(* IEC 61131-3 sources: plc-st-coding-agent/progress/evidence/f14_v10_full_20261113/jobs/codex_deepseek-v4pro (part 2) *)

(* ---- public-medium-05.candidate_02.st ---- *)
FUNCTION_BLOCK ProductionLineControl
(*
ENGINEERING_CONTRACT
MotorForward (PUB006/PUB007): manual ForwardButton iff not ReverseButton; auto hold while AutoStep=1 or AutoStep=3; deactivate at destination sensor B/C or on manual release/non-auto; simultaneous Forward/Reverse gives no motion.
MotorReverse (PUB004): manual ReverseButton iff not ForwardButton.
CompletionLight (PUB008): auto activate when C is reached and SensorC and ButtonC are TRUE, including same-scan arrival; retain while SensorC TRUE; reset only when SensorC FALSE.
AutoStep retains sequence state across scans; BOOL buttons are level-gated, no unstated edges.
*)
(* CONTRACT_RULES [] *)
VAR_INPUT
    Mode : BOOL;
    ForwardButton : BOOL;
    ReverseButton : BOOL;
    SensorA : BOOL;
    SensorB : BOOL;
    SensorC : BOOL;
    ButtonA : BOOL;
    ButtonB : BOOL;
    ButtonC : BOOL;
END_VAR
VAR_OUTPUT
    MotorForward : BOOL;
    MotorReverse : BOOL;
    CompletionLight : BOOL;
END_VAR
VAR
    AutoStep : INT := 0;
END_VAR

MotorForward := FALSE;
MotorReverse := FALSE;

IF NOT SensorC THEN
    CompletionLight := FALSE;
END_IF;

IF Mode THEN
    CASE AutoStep OF
        0:
            IF SensorA AND ButtonA THEN
                AutoStep := 1;
                MotorForward := TRUE;
            END_IF;

        1:
            IF SensorB THEN
                IF ButtonB THEN
                    AutoStep := 3;
                    MotorForward := TRUE;
                ELSE
                    AutoStep := 2;
                END_IF;
            ELSE
                MotorForward := TRUE;
            END_IF;

        2:
            IF ButtonB THEN
                AutoStep := 3;
                MotorForward := TRUE;
            END_IF;

        3:
            IF SensorC THEN
                AutoStep := 4;
                IF ButtonC THEN
                    CompletionLight := TRUE;
                END_IF;
            ELSE
                MotorForward := TRUE;
            END_IF;

        4:
            IF SensorC AND ButtonC THEN
                CompletionLight := TRUE;
            END_IF;
            IF NOT SensorC THEN
                AutoStep := 0;
            END_IF;
    END_CASE;
ELSE
    MotorForward := ForwardButton AND NOT ReverseButton;
    MotorReverse := ReverseButton AND NOT ForwardButton;
END_IF;
END_FUNCTION_BLOCK

(* ---- public-medium-05.candidate_03.st ---- *)
FUNCTION_BLOCK ProductionLineControl
(*
ENGINEERING_CONTRACT
MotorForward (PUB006/PUB007): manual ForwardButton iff not ReverseButton; auto hold while AutoStep=1 or AutoStep=3; deactivate at destination sensor B/C or on manual release/non-auto; simultaneous Forward/Reverse gives no motion.
MotorReverse (PUB004): manual ReverseButton iff not ForwardButton.
CompletionLight (PUB008): auto activate when C is reached and SensorC and ButtonC are TRUE, including same-scan arrival; retain while SensorC TRUE; reset only when SensorC FALSE.
AutoStep retains sequence state across scans; BOOL buttons are level-gated, no unstated edges.
*)
(* CONTRACT_RULES [] *)
VAR_INPUT
    Mode : BOOL;
    ForwardButton : BOOL;
    ReverseButton : BOOL;
    SensorA : BOOL;
    SensorB : BOOL;
    SensorC : BOOL;
    ButtonA : BOOL;
    ButtonB : BOOL;
    ButtonC : BOOL;
END_VAR
VAR_OUTPUT
    MotorForward : BOOL;
    MotorReverse : BOOL;
    CompletionLight : BOOL;
END_VAR
VAR
    AutoStep : INT := 0;
END_VAR

MotorForward := FALSE;
MotorReverse := FALSE;

IF NOT SensorC THEN
    CompletionLight := FALSE;
END_IF;

IF Mode THEN
    CASE AutoStep OF
        0:
            IF SensorA AND ButtonA THEN
                AutoStep := 1;
                MotorForward := TRUE;
            END_IF;

        1:
            IF SensorB THEN
                IF ButtonB THEN
                    AutoStep := 3;
                    MotorForward := TRUE;
                ELSE
                    AutoStep := 2;
                END_IF;
            ELSE
                MotorForward := TRUE;
            END_IF;

        2:
            IF ButtonB THEN
                AutoStep := 3;
                MotorForward := TRUE;
            END_IF;

        3:
            IF SensorC THEN
                AutoStep := 4;
                IF ButtonC THEN
                    CompletionLight := TRUE;
                END_IF;
            ELSE
                MotorForward := TRUE;
            END_IF;

        4:
            IF SensorC AND (CompletionLight OR ButtonC) THEN
                CompletionLight := TRUE;
            END_IF;
            IF NOT SensorC THEN
                AutoStep := 0;
            END_IF;
    END_CASE;
ELSE
    MotorForward := ForwardButton AND NOT ReverseButton;
    MotorReverse := ReverseButton AND NOT ForwardButton;
END_IF;
END_FUNCTION_BLOCK

(* ---- public-medium-05.raw_candidate_01.st ---- *)
FUNCTION_BLOCK ProductionLineControl
(*
ENGINEERING_CONTRACT
MotorForward (PUB001/PUB002/PUB003): activate manual ForwardButton or auto transfer state; hold through transfer to destination sensor; deactivate at destination sensor, manual release, or not in transfer state; simultaneous manual Forward/Reverse is interlocked, no motion.
MotorReverse (PUB002): activate only manual ReverseButton; no hold; deactivate on release or ForwardButton.
CompletionLight (PUB003): activate in auto at C while SensorC and ButtonC are TRUE; retain while SensorC remains TRUE; deactivation only when SensorC becomes FALSE; manual Mode does not reset it.
Bounds/units: BOOL inputs, BOOL outputs, discrete scan steps; buttons are level-gated, not edge-only.
Unspecified: simultaneous manual Forward/Reverse means no motion; automatic step is retained across mode changes.
*)
(* CONTRACT_RULES [] *)
VAR_INPUT
    Mode : BOOL;
    ForwardButton : BOOL;
    ReverseButton : BOOL;
    SensorA : BOOL;
    SensorB : BOOL;
    SensorC : BOOL;
    ButtonA : BOOL;
    ButtonB : BOOL;
    ButtonC : BOOL;
END_VAR
VAR_OUTPUT
    MotorForward : BOOL;
    MotorReverse : BOOL;
    CompletionLight : BOOL;
END_VAR
VAR
    AutoStep : INT := 0;
END_VAR

MotorForward := FALSE;
MotorReverse := FALSE;

IF NOT SensorC THEN
    CompletionLight := FALSE;
END_IF;

IF Mode THEN
    CASE AutoStep OF
        0:
            IF SensorA AND ButtonA THEN
                AutoStep := 1;
                MotorForward := TRUE;
            END_IF;

        1:
            IF SensorB THEN
                AutoStep := 2;
            END_IF;

        2:
            IF ButtonB THEN
                AutoStep := 3;
                MotorForward := TRUE;
            END_IF;

        3:
            IF SensorC THEN
                AutoStep := 4;
            END_IF;

        4:
            IF SensorC AND ButtonC THEN
                CompletionLight := TRUE;
            END_IF;
            IF NOT SensorC THEN
                AutoStep := 0;
            END_IF;
    END_CASE;
ELSE
    MotorForward := ForwardButton AND NOT ReverseButton;
    MotorReverse := ReverseButton AND NOT ForwardButton;
END_IF;
END_FUNCTION_BLOCK

(* ---- public-medium-05.raw_candidate_02.st ---- *)
FUNCTION_BLOCK ProductionLineControl
(*
ENGINEERING_CONTRACT
MotorForward (PUB006/PUB007): manual ForwardButton iff not ReverseButton; auto hold while AutoStep=1 or AutoStep=3; deactivate at destination sensor B/C or on manual release/non-auto; simultaneous Forward/Reverse gives no motion.
MotorReverse (PUB004): manual ReverseButton iff not ForwardButton.
CompletionLight (PUB008): auto activate when C is reached and SensorC and ButtonC are TRUE, including same-scan arrival; retain while SensorC TRUE; reset only when SensorC FALSE.
AutoStep retains sequence state across scans; BOOL buttons are level-gated, no unstated edges.
*)
(* CONTRACT_RULES [] *)
VAR_INPUT
    Mode : BOOL;
    ForwardButton : BOOL;
    ReverseButton : BOOL;
    SensorA : BOOL;
    SensorB : BOOL;
    SensorC : BOOL;
    ButtonA : BOOL;
    ButtonB : BOOL;
    ButtonC : BOOL;
END_VAR
VAR_OUTPUT
    MotorForward : BOOL;
    MotorReverse : BOOL;
    CompletionLight : BOOL;
END_VAR
VAR
    AutoStep : INT := 0;
END_VAR

MotorForward := FALSE;
MotorReverse := FALSE;

IF NOT SensorC THEN
    CompletionLight := FALSE;
END_IF;

IF Mode THEN
    CASE AutoStep OF
        0:
            IF SensorA AND ButtonA THEN
                AutoStep := 1;
                MotorForward := TRUE;
            END_IF;

        1:
            IF SensorB THEN
                IF ButtonB THEN
                    AutoStep := 3;
                    MotorForward := TRUE;
                ELSE
                    AutoStep := 2;
                END_IF;
            ELSE
                MotorForward := TRUE;
            END_IF;

        2:
            IF ButtonB THEN
                AutoStep := 3;
                MotorForward := TRUE;
            END_IF;

        3:
            IF SensorC THEN
                AutoStep := 4;
                IF ButtonC THEN
                    CompletionLight := TRUE;
                END_IF;
            ELSE
                MotorForward := TRUE;
            END_IF;

        4:
            IF SensorC AND ButtonC THEN
                CompletionLight := TRUE;
            END_IF;
            IF NOT SensorC THEN
                AutoStep := 0;
            END_IF;
    END_CASE;
ELSE
    MotorForward := ForwardButton AND NOT ReverseButton;
    MotorReverse := ReverseButton AND NOT ForwardButton;
END_IF;
END_FUNCTION_BLOCK

(* ---- public-medium-05.raw_candidate_03.st ---- *)
FUNCTION_BLOCK ProductionLineControl
(*
ENGINEERING_CONTRACT
MotorForward (PUB006/PUB007): manual ForwardButton iff not ReverseButton; auto hold while AutoStep=1 or AutoStep=3; deactivate at destination sensor B/C or on manual release/non-auto; simultaneous Forward/Reverse gives no motion.
MotorReverse (PUB004): manual ReverseButton iff not ForwardButton.
CompletionLight (PUB008): auto activate when C is reached and SensorC and ButtonC are TRUE, including same-scan arrival; retain while SensorC TRUE; reset only when SensorC FALSE.
AutoStep retains sequence state across scans; BOOL buttons are level-gated, no unstated edges.
*)
(* CONTRACT_RULES [] *)
VAR_INPUT
    Mode : BOOL;
    ForwardButton : BOOL;
    ReverseButton : BOOL;
    SensorA : BOOL;
    SensorB : BOOL;
    SensorC : BOOL;
    ButtonA : BOOL;
    ButtonB : BOOL;
    ButtonC : BOOL;
END_VAR
VAR_OUTPUT
    MotorForward : BOOL;
    MotorReverse : BOOL;
    CompletionLight : BOOL;
END_VAR
VAR
    AutoStep : INT := 0;
END_VAR

MotorForward := FALSE;
MotorReverse := FALSE;

IF NOT SensorC THEN
    CompletionLight := FALSE;
END_IF;

IF Mode THEN
    CASE AutoStep OF
        0:
            IF SensorA AND ButtonA THEN
                AutoStep := 1;
                MotorForward := TRUE;
            END_IF;

        1:
            IF SensorB THEN
                IF ButtonB THEN
                    AutoStep := 3;
                    MotorForward := TRUE;
                ELSE
                    AutoStep := 2;
                END_IF;
            ELSE
                MotorForward := TRUE;
            END_IF;

        2:
            IF ButtonB THEN
                AutoStep := 3;
                MotorForward := TRUE;
            END_IF;

        3:
            IF SensorC THEN
                AutoStep := 4;
                IF ButtonC THEN
                    CompletionLight := TRUE;
                END_IF;
            ELSE
                MotorForward := TRUE;
            END_IF;

        4:
            IF SensorC AND (CompletionLight OR ButtonC) THEN
                CompletionLight := TRUE;
            END_IF;
            IF NOT SensorC THEN
                AutoStep := 0;
            END_IF;
    END_CASE;
ELSE
    MotorForward := ForwardButton AND NOT ReverseButton;
    MotorReverse := ReverseButton AND NOT ForwardButton;
END_IF;
END_FUNCTION_BLOCK

(* ---- public-medium-06.candidate_01.st ---- *)
FUNCTION_BLOCK SlabThicknessMonitor
VAR_INPUT
    THICKNESS_FAULT : BOOL;
    THICKNESS_SIGNAL_VALID : BOOL;
    CUTTING_RUN : BOOL;
    FaultTimestamp : DINT;
    CycleTime : TIME;
END_VAR
VAR_OUTPUT
    THICKNESS_ALARM : BOOL;
    Slab_Fault_Counter : UINT;
    Slab_Runtime_Accumulator : LTIME;
    Slab_Fault_History : ARRAY[0..4] OF DINT;
END_VAR
VAR
    tmp_ValidFault : BOOL := FALSE;
    tmp_PrevValidFault : BOOL := FALSE;
    tmp_FaultRisingEdge : BOOL := FALSE;
    tmp_HoldRemaining : TIME := T#0MS;
    tmp_Initialized : BOOL := FALSE;
    tmp_Index : INT := 0;
    tmp_CycleLT : LTIME := LTIME#0S;
END_VAR

(* ENGINEERING_CONTRACT
- THICKNESS_ALARM: active immediately on valid fault true; held for >= 500 ms from each valid fault rising edge; remains active while fault persists; cleared on signal invalid or power-up. Signal invalid has priority over fault. PUB001/PUB004.
- Slab_Fault_Counter: increments on each FALSE-to-TRUE transition of the valid fault composite signal; persists across scans while signal invalid; UINT overflow is unspecified. PUB002/PUB004.
- Slab_Fault_History: index 0 is newest, older fault timestamps shift toward index 4 before overwriting; zero-filled on power-up and with no records. PUB002/PUB005.
- Slab_Runtime_Accumulator: adds TIME_TO_LTIME(CycleTime) only when signal valid, CUTTING_RUN is TRUE, and no thickness fault is present; otherwise value is retained. PUB003.
- Hold timing: timer set on the fault rising edge and decremented by CycleTime only on subsequent valid invocations; first satisfying hold interval is 500 ms. PUB001.
- Invalid signal: alarm and hold state are cleared; no fault record or runtime accumulation occurs. PUB004/PUB005.
*)
(* CONTRACT_RULES [] *)

IF NOT tmp_Initialized THEN
    THICKNESS_ALARM := FALSE;
    Slab_Fault_Counter := 0;
    Slab_Runtime_Accumulator := LTIME#0S;
    FOR tmp_Index := 0 TO 4 DO
        Slab_Fault_History[tmp_Index] := 0;
    END_FOR;
    tmp_HoldRemaining := T#0MS;
    tmp_PrevValidFault := FALSE;
    tmp_Initialized := TRUE;
END_IF;

tmp_ValidFault := THICKNESS_SIGNAL_VALID AND THICKNESS_FAULT;
tmp_FaultRisingEdge := tmp_ValidFault AND NOT tmp_PrevValidFault;

IF NOT THICKNESS_SIGNAL_VALID THEN
    THICKNESS_ALARM := FALSE;
    tmp_HoldRemaining := T#0MS;
ELSE
    IF tmp_FaultRisingEdge THEN
        Slab_Fault_Counter := Slab_Fault_Counter + 1;
        FOR tmp_Index := 4 TO 1 BY -1 DO
            Slab_Fault_History[tmp_Index] := Slab_Fault_History[tmp_Index - 1];
        END_FOR;
        Slab_Fault_History[0] := FaultTimestamp;
        tmp_HoldRemaining := T#500MS;
    ELSIF tmp_HoldRemaining > T#0MS THEN
        IF CycleTime > T#0MS THEN
            IF tmp_HoldRemaining >= CycleTime THEN
                tmp_HoldRemaining := tmp_HoldRemaining - CycleTime;
            ELSE
                tmp_HoldRemaining := T#0MS;
            END_IF;
        END_IF;
    END_IF;

    IF THICKNESS_FAULT OR (tmp_HoldRemaining > T#0MS) THEN
        THICKNESS_ALARM := TRUE;
    ELSE
        THICKNESS_ALARM := FALSE;
    END_IF;

    IF CUTTING_RUN AND NOT THICKNESS_FAULT AND (CycleTime > T#0MS) THEN
        tmp_CycleLT := TIME_TO_LTIME(CycleTime);
        Slab_Runtime_Accumulator := Slab_Runtime_Accumulator + tmp_CycleLT;
    END_IF;
END_IF;

tmp_PrevValidFault := tmp_ValidFault;
END_FUNCTION_BLOCK

(* ---- public-medium-06.raw_candidate_01.st ---- *)
FUNCTION_BLOCK SlabThicknessMonitor
VAR_INPUT
    THICKNESS_FAULT : BOOL;
    THICKNESS_SIGNAL_VALID : BOOL;
    CUTTING_RUN : BOOL;
    FaultTimestamp : DINT;
    CycleTime : TIME;
END_VAR
VAR_OUTPUT
    THICKNESS_ALARM : BOOL;
    Slab_Fault_Counter : UINT;
    Slab_Runtime_Accumulator : LTIME;
    Slab_Fault_History : ARRAY[0..4] OF DINT;
END_VAR
VAR
    tmp_ValidFault : BOOL := FALSE;
    tmp_PrevValidFault : BOOL := FALSE;
    tmp_FaultRisingEdge : BOOL := FALSE;
    tmp_HoldRemaining : TIME := T#0MS;
    tmp_Initialized : BOOL := FALSE;
    tmp_Index : INT := 0;
    tmp_CycleLT : LTIME := LTIME#0S;
END_VAR

(* ENGINEERING_CONTRACT
- THICKNESS_ALARM: active immediately on valid fault true; held for >= 500 ms from each valid fault rising edge; remains active while fault persists; cleared on signal invalid or power-up. Signal invalid has priority over fault. PUB001/PUB004.
- Slab_Fault_Counter: increments on each FALSE-to-TRUE transition of the valid fault composite signal; persists across scans while signal invalid; UINT overflow is unspecified. PUB002/PUB004.
- Slab_Fault_History: index 0 is newest, older fault timestamps shift toward index 4 before overwriting; zero-filled on power-up and with no records. PUB002/PUB005.
- Slab_Runtime_Accumulator: adds TIME_TO_LTIME(CycleTime) only when signal valid, CUTTING_RUN is TRUE, and no thickness fault is present; otherwise value is retained. PUB003.
- Hold timing: timer set on the fault rising edge and decremented by CycleTime only on subsequent valid invocations; first satisfying hold interval is 500 ms. PUB001.
- Invalid signal: alarm and hold state are cleared; no fault record or runtime accumulation occurs. PUB004/PUB005.
*)
(* CONTRACT_RULES [] *)

IF NOT tmp_Initialized THEN
    THICKNESS_ALARM := FALSE;
    Slab_Fault_Counter := 0;
    Slab_Runtime_Accumulator := LTIME#0S;
    FOR tmp_Index := 0 TO 4 DO
        Slab_Fault_History[tmp_Index] := 0;
    END_FOR;
    tmp_HoldRemaining := T#0MS;
    tmp_PrevValidFault := FALSE;
    tmp_Initialized := TRUE;
END_IF;

tmp_ValidFault := THICKNESS_SIGNAL_VALID AND THICKNESS_FAULT;
tmp_FaultRisingEdge := tmp_ValidFault AND NOT tmp_PrevValidFault;

IF NOT THICKNESS_SIGNAL_VALID THEN
    THICKNESS_ALARM := FALSE;
    tmp_HoldRemaining := T#0MS;
ELSE
    IF tmp_FaultRisingEdge THEN
        Slab_Fault_Counter := Slab_Fault_Counter + 1;
        FOR tmp_Index := 4 TO 1 BY -1 DO
            Slab_Fault_History[tmp_Index] := Slab_Fault_History[tmp_Index - 1];
        END_FOR;
        Slab_Fault_History[0] := FaultTimestamp;
        tmp_HoldRemaining := T#500MS;
    ELSIF tmp_HoldRemaining > T#0MS THEN
        IF CycleTime > T#0MS THEN
            IF tmp_HoldRemaining >= CycleTime THEN
                tmp_HoldRemaining := tmp_HoldRemaining - CycleTime;
            ELSE
                tmp_HoldRemaining := T#0MS;
            END_IF;
        END_IF;
    END_IF;

    IF THICKNESS_FAULT OR (tmp_HoldRemaining > T#0MS) THEN
        THICKNESS_ALARM := TRUE;
    ELSE
        THICKNESS_ALARM := FALSE;
    END_IF;

    IF CUTTING_RUN AND NOT THICKNESS_FAULT AND (CycleTime > T#0MS) THEN
        tmp_CycleLT := TIME_TO_LTIME(CycleTime);
        Slab_Runtime_Accumulator := Slab_Runtime_Accumulator + tmp_CycleLT;
    END_IF;
END_IF;

tmp_PrevValidFault := tmp_ValidFault;
END_FUNCTION_BLOCK

(* ---- public-medium-07.candidate_01.st ---- *)
(* ENGINEERING_CONTRACT
 * SUPPLY_FAN_RUN: activation requires OCCUPANCY_DETECTED=TRUE and selector <> 3
 * continuously for T#30S; holds while those conditions remain; occupancy loss or Night
 * deactivates immediately, resets timer, and recovery requires full T#30S (PUB002, PUB007).
 * TEMP_SETPOINT_ADJUST: recomputed every scan from current occupancy, energy-saving state
 * and HVAC mode; no latch or extra hold beyond current inputs (PUB003, PUB004, PUB005).
 * Same-scan priority: timer-enable is computed before TON, then fan Q and adjustment update
 * in the same scan; no edge-only triggers or resets beyond stated conditions.
 * Units/bounds: delay is exact T#30S; adjustment is integral degC clamped to [-4,4];
 * power-up outputs initialize to FALSE/OFF and 0 under standard VAR defaults (PUB006).
 *)
(* CONTRACT_RULES [] *)
FUNCTION_BLOCK FB_OfficeHvacControl
VAR_INPUT
    OCCUPANCY_DETECTED : BOOL;
    ENERGY_SAVING_MODE : BOOL;
    HVAC_MODE_SELECTOR : INT;
END_VAR
VAR_OUTPUT
    SUPPLY_FAN_RUN : BOOL;
    TEMP_SETPOINT_ADJUST : INT;
END_VAR
VAR
    fanTimer : TON;
    tmp_FanEnable : BOOL;
END_VAR

tmp_FanEnable := OCCUPANCY_DETECTED AND (HVAC_MODE_SELECTOR <> 3);

fanTimer(IN := tmp_FanEnable, PT := T#30S);
SUPPLY_FAN_RUN := fanTimer.Q;

CASE HVAC_MODE_SELECTOR OF
    0:
        IF OCCUPANCY_DETECTED THEN
            TEMP_SETPOINT_ADJUST := 0;
        ELSIF ENERGY_SAVING_MODE THEN
            TEMP_SETPOINT_ADJUST := 3;
        ELSE
            TEMP_SETPOINT_ADJUST := 2;
        END_IF;
    1:
        IF OCCUPANCY_DETECTED THEN
            TEMP_SETPOINT_ADJUST := 0;
        ELSE
            TEMP_SETPOINT_ADJUST := 1;
        END_IF;
    2:
        IF OCCUPANCY_DETECTED THEN
            TEMP_SETPOINT_ADJUST := 0;
        ELSE
            TEMP_SETPOINT_ADJUST := 4;
        END_IF;
    3:
        TEMP_SETPOINT_ADJUST := 4;
    ELSE
        TEMP_SETPOINT_ADJUST := 0;
END_CASE;

IF TEMP_SETPOINT_ADJUST < -4 THEN
    TEMP_SETPOINT_ADJUST := -4;
ELSIF TEMP_SETPOINT_ADJUST > 4 THEN
    TEMP_SETPOINT_ADJUST := 4;
END_IF;

END_FUNCTION_BLOCK

(* ---- public-medium-07.raw_candidate_01.st ---- *)
(* ENGINEERING_CONTRACT
 * SUPPLY_FAN_RUN: activation requires OCCUPANCY_DETECTED=TRUE and selector <> 3
 * continuously for T#30S; holds while those conditions remain; occupancy loss or Night
 * deactivates immediately, resets timer, and recovery requires full T#30S (PUB002, PUB007).
 * TEMP_SETPOINT_ADJUST: recomputed every scan from current occupancy, energy-saving state
 * and HVAC mode; no latch or extra hold beyond current inputs (PUB003, PUB004, PUB005).
 * Same-scan priority: timer-enable is computed before TON, then fan Q and adjustment update
 * in the same scan; no edge-only triggers or resets beyond stated conditions.
 * Units/bounds: delay is exact T#30S; adjustment is integral degC clamped to [-4,4];
 * power-up outputs initialize to FALSE/OFF and 0 under standard VAR defaults (PUB006).
 *)
(* CONTRACT_RULES [] *)
FUNCTION_BLOCK FB_OfficeHvacControl
VAR_INPUT
    OCCUPANCY_DETECTED : BOOL;
    ENERGY_SAVING_MODE : BOOL;
    HVAC_MODE_SELECTOR : INT;
END_VAR
VAR_OUTPUT
    SUPPLY_FAN_RUN : BOOL;
    TEMP_SETPOINT_ADJUST : INT;
END_VAR
VAR
    fanTimer : TON;
    tmp_FanEnable : BOOL;
END_VAR

tmp_FanEnable := OCCUPANCY_DETECTED AND (HVAC_MODE_SELECTOR <> 3);

fanTimer(IN := tmp_FanEnable, PT := T#30S);
SUPPLY_FAN_RUN := fanTimer.Q;

CASE HVAC_MODE_SELECTOR OF
    0:
        IF OCCUPANCY_DETECTED THEN
            TEMP_SETPOINT_ADJUST := 0;
        ELSIF ENERGY_SAVING_MODE THEN
            TEMP_SETPOINT_ADJUST := 3;
        ELSE
            TEMP_SETPOINT_ADJUST := 2;
        END_IF;
    1:
        IF OCCUPANCY_DETECTED THEN
            TEMP_SETPOINT_ADJUST := 0;
        ELSE
            TEMP_SETPOINT_ADJUST := 1;
        END_IF;
    2:
        IF OCCUPANCY_DETECTED THEN
            TEMP_SETPOINT_ADJUST := 0;
        ELSE
            TEMP_SETPOINT_ADJUST := 4;
        END_IF;
    3:
        TEMP_SETPOINT_ADJUST := 4;
    ELSE
        TEMP_SETPOINT_ADJUST := 0;
END_CASE;

IF TEMP_SETPOINT_ADJUST < -4 THEN
    TEMP_SETPOINT_ADJUST := -4;
ELSIF TEMP_SETPOINT_ADJUST > 4 THEN
    TEMP_SETPOINT_ADJUST := 4;
END_IF;

END_FUNCTION_BLOCK

(* ---- public-medium-08.candidate_01.st ---- *)
(* ENGINEERING_CONTRACT
- ipValue is recomputed from ipText on every scan; no retention/latch.
- Valid: exactly four nonempty all-digit segments, each value 0..255 inclusive.
- Network byte order: first segment is MSB, fourth segment is LSB.
- Malformed text, nondigit, empty segment, wrong segment count, or out-of-range
  value sets ipValue := 0 in that same scan.
- 0.0.0.0 is valid and produces 0.
- Leading zeros are accepted as decimal digits; their rejection is unspecified.
- Invalid-input returns leave ipValue at its preassigned value of 0.
*)
(* CONTRACT_RULES [] *)
FUNCTION_BLOCK FB_IPv4Parser
VAR_INPUT
    ipText : STRING(254);
END_VAR
VAR_OUTPUT
    ipValue : UDINT;
END_VAR
VAR
    tmp_Length : INT;
    tmp_Pos : INT;
    tmp_SegmentCount : INT;
    tmp_DigitCount : INT;
    tmp_SegmentValue : UDINT;
    tmp_CharCode : UDINT;
END_VAR

ipValue := 0;
tmp_Length := LEN(ipText);
tmp_Pos := 0;
tmp_SegmentCount := 0;
tmp_DigitCount := 0;
tmp_SegmentValue := 0;
tmp_CharCode := 0;

IF tmp_Length <= 0 THEN
    RETURN;
END_IF;

WHILE tmp_Pos < tmp_Length DO
    tmp_CharCode := BYTE_TO_UDINT(ipText[tmp_Pos]);

    IF (tmp_CharCode >= 48) AND (tmp_CharCode <= 57) THEN
        tmp_DigitCount := tmp_DigitCount + 1;
        tmp_SegmentValue := (tmp_SegmentValue * 10) + (tmp_CharCode - 48);

        IF tmp_SegmentValue > 255 THEN
            RETURN;
        END_IF;
    ELSIF tmp_CharCode = 46 THEN
        IF tmp_DigitCount <= 0 THEN
            RETURN;
        END_IF;

        tmp_SegmentCount := tmp_SegmentCount + 1;

        IF tmp_SegmentCount >= 4 THEN
            RETURN;
        END_IF;

        ipValue := (SHL(ipValue, 8)) OR tmp_SegmentValue;
        tmp_SegmentValue := 0;
        tmp_DigitCount := 0;
    ELSE
        RETURN;
    END_IF;

    tmp_Pos := tmp_Pos + 1;
END_WHILE;

IF tmp_DigitCount <= 0 THEN
    RETURN;
END_IF;

tmp_SegmentCount := tmp_SegmentCount + 1;

IF tmp_SegmentCount <> 4 THEN
    RETURN;
END_IF;

ipValue := (SHL(ipValue, 8)) OR tmp_SegmentValue;

END_FUNCTION_BLOCK

(* ---- public-medium-08.candidate_02.st ---- *)
(* ENGINEERING_CONTRACT
- ipValue is recomputed from ipText on every scan; no retention/latch.
- Valid: exactly four nonempty all-digit segments, each value 0..255 inclusive.
- Network byte order: first segment is MSB, fourth segment is LSB.
- Malformed text, nondigit, empty segment, wrong segment count, or out-of-range
  value sets ipValue := 0 in that same scan.
- 0.0.0.0 is valid and produces 0.
- Leading zeros are accepted as decimal digits; their rejection is unspecified.
- Invalid-input returns leave ipValue at its preassigned value of 0.
*)
(* CONTRACT_RULES [] *)
FUNCTION_BLOCK FB_IPv4Parser
VAR_INPUT
    ipText : STRING(254);
END_VAR
VAR_OUTPUT
    ipValue : UDINT;
END_VAR
VAR
    tmp_Length : INT;
    tmp_Pos : INT;
    tmp_SegmentCount : INT;
    tmp_DigitCount : INT;
    tmp_SegmentValue : UDINT;
    tmp_CharCode : UDINT;
    tmp_Accum : UDINT;
END_VAR

ipValue := 0;
tmp_Accum := 0;
tmp_Length := LEN(ipText);
tmp_Pos := 0;
tmp_SegmentCount := 0;
tmp_DigitCount := 0;
tmp_SegmentValue := 0;
tmp_CharCode := 0;

IF tmp_Length <= 0 THEN
    RETURN;
END_IF;

WHILE tmp_Pos < tmp_Length DO
    tmp_CharCode := BYTE_TO_UDINT(ipText[tmp_Pos]);

    IF (tmp_CharCode >= 48) AND (tmp_CharCode <= 57) THEN
        tmp_DigitCount := tmp_DigitCount + 1;
        tmp_SegmentValue := (tmp_SegmentValue * 10) + (tmp_CharCode - 48);

        IF tmp_SegmentValue > 255 THEN
            RETURN;
        END_IF;
    ELSIF tmp_CharCode = 46 THEN
        IF tmp_DigitCount <= 0 THEN
            RETURN;
        END_IF;

        tmp_SegmentCount := tmp_SegmentCount + 1;

        IF tmp_SegmentCount >= 4 THEN
            RETURN;
        END_IF;

        tmp_Accum := (SHL(tmp_Accum, 8)) OR tmp_SegmentValue;
        tmp_SegmentValue := 0;
        tmp_DigitCount := 0;
    ELSE
        RETURN;
    END_IF;

    tmp_Pos := tmp_Pos + 1;
END_WHILE;

IF tmp_DigitCount <= 0 THEN
    RETURN;
END_IF;

tmp_SegmentCount := tmp_SegmentCount + 1;

IF tmp_SegmentCount <> 4 THEN
    RETURN;
END_IF;

tmp_Accum := (SHL(tmp_Accum, 8)) OR tmp_SegmentValue;
ipValue := tmp_Accum;

END_FUNCTION_BLOCK

(* ---- public-medium-08.raw_candidate_01.st ---- *)
(* ENGINEERING_CONTRACT
- ipValue is recomputed from ipText on every scan; no retention/latch.
- Valid: exactly four nonempty all-digit segments, each value 0..255 inclusive.
- Network byte order: first segment is MSB, fourth segment is LSB.
- Malformed text, nondigit, empty segment, wrong segment count, or out-of-range
  value sets ipValue := 0 in that same scan.
- 0.0.0.0 is valid and produces 0.
- Leading zeros are accepted as decimal digits; their rejection is unspecified.
- Invalid-input returns leave ipValue at its preassigned value of 0.
*)
(* CONTRACT_RULES [] *)
FUNCTION_BLOCK FB_IPv4Parser
VAR_INPUT
    ipText : STRING(254);
END_VAR
VAR_OUTPUT
    ipValue : UDINT;
END_VAR
VAR
    tmp_Length : INT;
    tmp_Pos : INT;
    tmp_SegmentCount : INT;
    tmp_DigitCount : INT;
    tmp_SegmentValue : UDINT;
    tmp_CharCode : UDINT;
END_VAR

ipValue := 0;
tmp_Length := LEN(ipText);
tmp_Pos := 0;
tmp_SegmentCount := 0;
tmp_DigitCount := 0;
tmp_SegmentValue := 0;
tmp_CharCode := 0;

IF tmp_Length <= 0 THEN
    RETURN;
END_IF;

WHILE tmp_Pos < tmp_Length DO
    tmp_CharCode := BYTE_TO_UDINT(ipText[tmp_Pos]);

    IF (tmp_CharCode >= 48) AND (tmp_CharCode <= 57) THEN
        tmp_DigitCount := tmp_DigitCount + 1;
        tmp_SegmentValue := (tmp_SegmentValue * 10) + (tmp_CharCode - 48);

        IF tmp_SegmentValue > 255 THEN
            RETURN;
        END_IF;
    ELSIF tmp_CharCode = 46 THEN
        IF tmp_DigitCount <= 0 THEN
            RETURN;
        END_IF;

        tmp_SegmentCount := tmp_SegmentCount + 1;

        IF tmp_SegmentCount >= 4 THEN
            RETURN;
        END_IF;

        ipValue := (SHL(ipValue, 8)) OR tmp_SegmentValue;
        tmp_SegmentValue := 0;
        tmp_DigitCount := 0;
    ELSE
        RETURN;
    END_IF;

    tmp_Pos := tmp_Pos + 1;
END_WHILE;

IF tmp_DigitCount <= 0 THEN
    RETURN;
END_IF;

tmp_SegmentCount := tmp_SegmentCount + 1;

IF tmp_SegmentCount <> 4 THEN
    RETURN;
END_IF;

ipValue := (SHL(ipValue, 8)) OR tmp_SegmentValue;

END_FUNCTION_BLOCK

(* ---- public-medium-08.raw_candidate_02.st ---- *)
(* ENGINEERING_CONTRACT
- ipValue is recomputed from ipText on every scan; no retention/latch.
- Valid: exactly four nonempty all-digit segments, each value 0..255 inclusive.
- Network byte order: first segment is MSB, fourth segment is LSB.
- Malformed text, nondigit, empty segment, wrong segment count, or out-of-range
  value sets ipValue := 0 in that same scan.
- 0.0.0.0 is valid and produces 0.
- Leading zeros are accepted as decimal digits; their rejection is unspecified.
- Invalid-input returns leave ipValue at its preassigned value of 0.
*)
(* CONTRACT_RULES [] *)
FUNCTION_BLOCK FB_IPv4Parser
VAR_INPUT
    ipText : STRING(254);
END_VAR
VAR_OUTPUT
    ipValue : UDINT;
END_VAR
VAR
    tmp_Length : INT;
    tmp_Pos : INT;
    tmp_SegmentCount : INT;
    tmp_DigitCount : INT;
    tmp_SegmentValue : UDINT;
    tmp_CharCode : UDINT;
    tmp_Accum : UDINT;
END_VAR

ipValue := 0;
tmp_Accum := 0;
tmp_Length := LEN(ipText);
tmp_Pos := 0;
tmp_SegmentCount := 0;
tmp_DigitCount := 0;
tmp_SegmentValue := 0;
tmp_CharCode := 0;

IF tmp_Length <= 0 THEN
    RETURN;
END_IF;

WHILE tmp_Pos < tmp_Length DO
    tmp_CharCode := BYTE_TO_UDINT(ipText[tmp_Pos]);

    IF (tmp_CharCode >= 48) AND (tmp_CharCode <= 57) THEN
        tmp_DigitCount := tmp_DigitCount + 1;
        tmp_SegmentValue := (tmp_SegmentValue * 10) + (tmp_CharCode - 48);

        IF tmp_SegmentValue > 255 THEN
            RETURN;
        END_IF;
    ELSIF tmp_CharCode = 46 THEN
        IF tmp_DigitCount <= 0 THEN
            RETURN;
        END_IF;

        tmp_SegmentCount := tmp_SegmentCount + 1;

        IF tmp_SegmentCount >= 4 THEN
            RETURN;
        END_IF;

        tmp_Accum := (SHL(tmp_Accum, 8)) OR tmp_SegmentValue;
        tmp_SegmentValue := 0;
        tmp_DigitCount := 0;
    ELSE
        RETURN;
    END_IF;

    tmp_Pos := tmp_Pos + 1;
END_WHILE;

IF tmp_DigitCount <= 0 THEN
    RETURN;
END_IF;

tmp_SegmentCount := tmp_SegmentCount + 1;

IF tmp_SegmentCount <> 4 THEN
    RETURN;
END_IF;

tmp_Accum := (SHL(tmp_Accum, 8)) OR tmp_SegmentValue;
ipValue := tmp_Accum;

END_FUNCTION_BLOCK

(* ---- self-easy-01.candidate_01.st ---- *)
FUNCTION_BLOCK FB
VAR_INPUT
    enable : BOOL;
    values : ARRAY[1..8] OF INT;
    count : INT;
    avgEnable : BOOL;
END_VAR
VAR_OUTPUT
    avgOut : REAL;
END_VAR
VAR
    tmp_i : INT;
    tmp_len : INT;
    tmp_sum : LINT;
END_VAR

(* ENGINEERING_CONTRACT
- Writes avgOut only when enable=TRUE AND avgEnable=TRUE AND count>=1.
- Holds previous avgOut for !enable (PUB003), !avgEnable (PUB007), or count<=0 (PUB005).
- count>8 uses first 8 entries only; no out-of-range access (PUB006).
- Same-scan priority: hold condition is checked first, so no competing write occurs.
- Activation/deactivation: no reset input; output is replaced only by a valid calculation.
- Units/boundaries: avgOut REAL = LINT sum / REAL length; sum uses LINT (PUB008, PUB009).
*)

(* CONTRACT_RULES [] *)

IF enable AND avgEnable AND (count > 0) THEN
    IF count >= 8 THEN
        tmp_len := 8;
    ELSE
        tmp_len := count;
    END_IF;

    tmp_sum := 0;

    FOR tmp_i := 1 TO tmp_len DO
        tmp_sum := tmp_sum + INT_TO_LINT(values[tmp_i]);
    END_FOR;

    avgOut := LINT_TO_REAL(tmp_sum) / INT_TO_REAL(tmp_len);
END_IF;

END_FUNCTION_BLOCK

(* ---- self-easy-01.raw_candidate_01.st ---- *)
FUNCTION_BLOCK FB
VAR_INPUT
    enable : BOOL;
    values : ARRAY[1..8] OF INT;
    count : INT;
    avgEnable : BOOL;
END_VAR
VAR_OUTPUT
    avgOut : REAL;
END_VAR
VAR
    tmp_i : INT;
    tmp_len : INT;
    tmp_sum : LINT;
END_VAR

(* ENGINEERING_CONTRACT
- Writes avgOut only when enable=TRUE AND avgEnable=TRUE AND count>=1.
- Holds previous avgOut for !enable (PUB003), !avgEnable (PUB007), or count<=0 (PUB005).
- count>8 uses first 8 entries only; no out-of-range access (PUB006).
- Same-scan priority: hold condition is checked first, so no competing write occurs.
- Activation/deactivation: no reset input; output is replaced only by a valid calculation.
- Units/boundaries: avgOut REAL = LINT sum / REAL length; sum uses LINT (PUB008, PUB009).
*)

(* CONTRACT_RULES [] *)

IF enable AND avgEnable AND (count > 0) THEN
    IF count >= 8 THEN
        tmp_len := 8;
    ELSE
        tmp_len := count;
    END_IF;

    tmp_sum := 0;

    FOR tmp_i := 1 TO tmp_len DO
        tmp_sum := tmp_sum + INT_TO_LINT(values[tmp_i]);
    END_FOR;

    avgOut := LINT_TO_REAL(tmp_sum) / INT_TO_REAL(tmp_len);
END_IF;

END_FUNCTION_BLOCK

(* ---- self-easy-02.candidate_01.st ---- *)
(*
ENGINEERING_CONTRACT
- alarmHigh: active if tankLevel >= 85.0; once active, retains until a rising resetBtn occurs while tankLevel < 85.0; danger on the same scan as reset wins.
- alarmLow: active if tankLevel <= 15.0; once active, retains until a rising resetBtn occurs while tankLevel > 15.0; danger on the same scan as reset wins.
- reset edge: rising only when resetBtn is TRUE and the stored previous value is FALSE; holding resetBtn generates no additional resets.
- pumpRun: evaluated after alarm updates, TRUE only when inletPermit, !alarmHigh, and !alarmLow.
- outletValveOpen: evaluated after alarm updates, equals !alarmLow.
- outletFlow: observation input only, not used.
- Units: tankLevel is REAL percent; thresholds are inclusive as stated.
*)
(* CONTRACT_RULES [] *)
FUNCTION_BLOCK FB
VAR_INPUT
    tankLevel : REAL;
    outletFlow : REAL;
    inletPermit : BOOL;
    resetBtn : BOOL;
END_VAR
VAR_OUTPUT
    pumpRun : BOOL;
    alarmHigh : BOOL;
    alarmLow : BOOL;
    outletValveOpen : BOOL;
END_VAR
VAR
    prevResetBtn : BOOL := FALSE;
    tmp_highDanger : BOOL;
    tmp_lowDanger : BOOL;
    tmp_resetRise : BOOL;
END_VAR

tmp_resetRise := resetBtn AND NOT prevResetBtn;

tmp_highDanger := tankLevel >= 85.0;
tmp_lowDanger := tankLevel <= 15.0;

alarmHigh := tmp_highDanger OR (alarmHigh AND NOT tmp_resetRise);
alarmLow := tmp_lowDanger OR (alarmLow AND NOT tmp_resetRise);

pumpRun := inletPermit AND NOT alarmHigh AND NOT alarmLow;
outletValveOpen := NOT alarmLow;

prevResetBtn := resetBtn;

END_FUNCTION_BLOCK

(* ---- self-easy-02.raw_candidate_01.st ---- *)
(*
ENGINEERING_CONTRACT
- alarmHigh: active if tankLevel >= 85.0; once active, retains until a rising resetBtn occurs while tankLevel < 85.0; danger on the same scan as reset wins.
- alarmLow: active if tankLevel <= 15.0; once active, retains until a rising resetBtn occurs while tankLevel > 15.0; danger on the same scan as reset wins.
- reset edge: rising only when resetBtn is TRUE and the stored previous value is FALSE; holding resetBtn generates no additional resets.
- pumpRun: evaluated after alarm updates, TRUE only when inletPermit, !alarmHigh, and !alarmLow.
- outletValveOpen: evaluated after alarm updates, equals !alarmLow.
- outletFlow: observation input only, not used.
- Units: tankLevel is REAL percent; thresholds are inclusive as stated.
*)
(* CONTRACT_RULES [] *)
FUNCTION_BLOCK FB
VAR_INPUT
    tankLevel : REAL;
    outletFlow : REAL;
    inletPermit : BOOL;
    resetBtn : BOOL;
END_VAR
VAR_OUTPUT
    pumpRun : BOOL;
    alarmHigh : BOOL;
    alarmLow : BOOL;
    outletValveOpen : BOOL;
END_VAR
VAR
    prevResetBtn : BOOL := FALSE;
    tmp_highDanger : BOOL;
    tmp_lowDanger : BOOL;
    tmp_resetRise : BOOL;
END_VAR

tmp_resetRise := resetBtn AND NOT prevResetBtn;

tmp_highDanger := tankLevel >= 85.0;
tmp_lowDanger := tankLevel <= 15.0;

alarmHigh := tmp_highDanger OR (alarmHigh AND NOT tmp_resetRise);
alarmLow := tmp_lowDanger OR (alarmLow AND NOT tmp_resetRise);

pumpRun := inletPermit AND NOT alarmHigh AND NOT alarmLow;
outletValveOpen := NOT alarmLow;

prevResetBtn := resetBtn;

END_FUNCTION_BLOCK

(* ---- self-hard-01.candidate_01.st ---- *)
(*
ENGINEERING_CONTRACT
alarmActive: set when flowLow is TRUE (PUB001); holds when flowLow clears unacknowledged (PUB002); clears on current rising ack with flowLow FALSE, or automatically after already acknowledged condition loss (PUB003, S6).
alarmAcked: cleared for an active unacknowledged condition; set by rising ack while flowLow remains TRUE, or when unacknowledged flowLow clears; cleared together with alarmActive on pending-clear ack (PUB002-PUB003, S7).
highHigh: equals NOT sensorOK every scan; no latch and no cross-suppression of alarmActive/alarmAcked (PUB004, S3, S5).
Same-scan priority: rising ack uses current ackBtn sample; flowLow/ack/sensorOK effects are independent; no hidden reset, timer, or extra edge trigger is added.
Units/bounds: all public values are BOOL per scan.
*)
(* CONTRACT_RULES [] *)
FUNCTION_BLOCK FB
VAR_INPUT
    flowLow : BOOL;
    ackBtn : BOOL;
    sensorOK : BOOL;
END_VAR
VAR_OUTPUT
    alarmActive : BOOL;
    alarmAcked : BOOL;
    highHigh : BOOL;
END_VAR
VAR
    local_prevAckBtn : BOOL := FALSE;
    local_prevFlowLow : BOOL := FALSE;
    local_prevAlarmActive : BOOL := FALSE;
    local_prevAlarmAcked : BOOL := FALSE;
    local_risingAck : BOOL;
    local_prevFlowAckedTerm : BOOL;
    local_prevRetainAckTerm : BOOL;
END_VAR

local_risingAck := ackBtn AND NOT local_prevAckBtn;

highHigh := NOT sensorOK;

local_prevFlowAckedTerm := local_prevFlowLow AND local_prevAlarmAcked;
alarmActive := flowLow OR (local_prevAlarmActive AND NOT local_risingAck AND NOT local_prevFlowAckedTerm);

local_prevRetainAckTerm := local_prevFlowLow AND local_prevAlarmActive AND local_prevAlarmAcked;
alarmAcked := alarmActive AND (NOT flowLow OR local_risingAck OR local_prevRetainAckTerm);

local_prevAckBtn := ackBtn;
local_prevFlowLow := flowLow;
local_prevAlarmActive := alarmActive;
local_prevAlarmAcked := alarmAcked;

(* ---- self-hard-01.candidate_02.st ---- *)
(*
ENGINEERING_CONTRACT
alarmActive: set when flowLow is TRUE (PUB001); holds when flowLow clears unacknowledged (PUB002); clears on current rising ack with flowLow FALSE, or automatically after already acknowledged condition loss (PUB003, S6).
alarmAcked: cleared for an active unacknowledged condition; set by rising ack while flowLow remains TRUE, or when unacknowledged flowLow clears; cleared together with alarmActive on pending-clear ack (PUB002-PUB003, S7).
highHigh: equals NOT sensorOK every scan; no latch and no cross-suppression of alarmActive/alarmAcked (PUB004, S3, S5).
Same-scan priority: rising ack uses current ackBtn sample; flowLow/ack/sensorOK effects are independent; no hidden reset, timer, or extra edge trigger is added.
Units/bounds: all public values are BOOL per scan.
*)
(* CONTRACT_RULES [] *)
FUNCTION_BLOCK FB
VAR_INPUT
    flowLow : BOOL;
    ackBtn : BOOL;
    sensorOK : BOOL;
END_VAR
VAR_OUTPUT
    alarmActive : BOOL;
    alarmAcked : BOOL;
    highHigh : BOOL;
END_VAR
VAR
    local_prevAckBtn : BOOL := FALSE;
    local_prevFlowLow : BOOL := FALSE;
    local_prevAlarmActive : BOOL := FALSE;
    local_prevAlarmAcked : BOOL := FALSE;
    local_risingAck : BOOL;
    local_prevFlowAckedTerm : BOOL;
    local_prevRetainAckTerm : BOOL;
END_VAR

local_risingAck := ackBtn AND NOT local_prevAckBtn;

highHigh := NOT sensorOK;

local_prevFlowAckedTerm := local_prevFlowLow AND local_prevAlarmAcked;
alarmActive := flowLow OR (local_prevAlarmActive AND NOT local_risingAck AND NOT local_prevFlowAckedTerm);

local_prevRetainAckTerm := local_prevFlowLow AND local_prevAlarmActive AND local_prevAlarmAcked;
alarmAcked := alarmActive AND (NOT flowLow OR local_risingAck OR local_prevRetainAckTerm);

local_prevAckBtn := ackBtn;
local_prevFlowLow := flowLow;
local_prevAlarmActive := alarmActive;
local_prevAlarmAcked := alarmAcked;

END_FUNCTION_BLOCK

(* ---- self-hard-01.raw_candidate_01.st ---- *)
(*
ENGINEERING_CONTRACT
alarmActive: set when flowLow is TRUE (PUB001); holds when flowLow clears unacknowledged (PUB002); clears on current rising ack with flowLow FALSE, or automatically after already acknowledged condition loss (PUB003, S6).
alarmAcked: cleared for an active unacknowledged condition; set by rising ack while flowLow remains TRUE, or when unacknowledged flowLow clears; cleared together with alarmActive on pending-clear ack (PUB002-PUB003, S7).
highHigh: equals NOT sensorOK every scan; no latch and no cross-suppression of alarmActive/alarmAcked (PUB004, S3, S5).
Same-scan priority: rising ack uses current ackBtn sample; flowLow/ack/sensorOK effects are independent; no hidden reset, timer, or extra edge trigger is added.
Units/bounds: all public values are BOOL per scan.
*)
(* CONTRACT_RULES [] *)
FUNCTION_BLOCK FB
VAR_INPUT
    flowLow : BOOL;
    ackBtn : BOOL;
    sensorOK : BOOL;
END_VAR
VAR_OUTPUT
    alarmActive : BOOL;
    alarmAcked : BOOL;
    highHigh : BOOL;
END_VAR
VAR
    local_prevAckBtn : BOOL := FALSE;
    local_prevFlowLow : BOOL := FALSE;
    local_prevAlarmActive : BOOL := FALSE;
    local_prevAlarmAcked : BOOL := FALSE;
    local_risingAck : BOOL;
    local_prevFlowAckedTerm : BOOL;
    local_prevRetainAckTerm : BOOL;
END_VAR

local_risingAck := ackBtn AND NOT local_prevAckBtn;

highHigh := NOT sensorOK;

local_prevFlowAckedTerm := local_prevFlowLow AND local_prevAlarmAcked;
alarmActive := flowLow OR (local_prevAlarmActive AND NOT local_risingAck AND NOT local_prevFlowAckedTerm);

local_prevRetainAckTerm := local_prevFlowLow AND local_prevAlarmActive AND local_prevAlarmAcked;
alarmAcked := alarmActive AND (NOT flowLow OR local_risingAck OR local_prevRetainAckTerm);

local_prevAckBtn := ackBtn;
local_prevFlowLow := flowLow;
local_prevAlarmActive := alarmActive;
local_prevAlarmAcked := alarmAcked;

(* ---- self-hard-01.raw_candidate_02.st ---- *)
(*
ENGINEERING_CONTRACT
alarmActive: set when flowLow is TRUE (PUB001); holds when flowLow clears unacknowledged (PUB002); clears on current rising ack with flowLow FALSE, or automatically after already acknowledged condition loss (PUB003, S6).
alarmAcked: cleared for an active unacknowledged condition; set by rising ack while flowLow remains TRUE, or when unacknowledged flowLow clears; cleared together with alarmActive on pending-clear ack (PUB002-PUB003, S7).
highHigh: equals NOT sensorOK every scan; no latch and no cross-suppression of alarmActive/alarmAcked (PUB004, S3, S5).
Same-scan priority: rising ack uses current ackBtn sample; flowLow/ack/sensorOK effects are independent; no hidden reset, timer, or extra edge trigger is added.
Units/bounds: all public values are BOOL per scan.
*)
(* CONTRACT_RULES [] *)
FUNCTION_BLOCK FB
VAR_INPUT
    flowLow : BOOL;
    ackBtn : BOOL;
    sensorOK : BOOL;
END_VAR
VAR_OUTPUT
    alarmActive : BOOL;
    alarmAcked : BOOL;
    highHigh : BOOL;
END_VAR
VAR
    local_prevAckBtn : BOOL := FALSE;
    local_prevFlowLow : BOOL := FALSE;
    local_prevAlarmActive : BOOL := FALSE;
    local_prevAlarmAcked : BOOL := FALSE;
    local_risingAck : BOOL;
    local_prevFlowAckedTerm : BOOL;
    local_prevRetainAckTerm : BOOL;
END_VAR

local_risingAck := ackBtn AND NOT local_prevAckBtn;

highHigh := NOT sensorOK;

local_prevFlowAckedTerm := local_prevFlowLow AND local_prevAlarmAcked;
alarmActive := flowLow OR (local_prevAlarmActive AND NOT local_risingAck AND NOT local_prevFlowAckedTerm);

local_prevRetainAckTerm := local_prevFlowLow AND local_prevAlarmActive AND local_prevAlarmAcked;
alarmAcked := alarmActive AND (NOT flowLow OR local_risingAck OR local_prevRetainAckTerm);

local_prevAckBtn := ackBtn;
local_prevFlowLow := flowLow;
local_prevAlarmActive := alarmActive;
local_prevAlarmAcked := alarmAcked;

END_FUNCTION_BLOCK

(* ---- self-hard-02.candidate_01.st ---- *)
FUNCTION_BLOCK FB
VAR_INPUT
    startBtn : BOOL;
    abortBtn : BOOL;
    setpoint : REAL;
    pv : REAL;
    maxDuration : INT;
END_VAR
VAR_OUTPUT
    elapsed : INT;
    phase : INT;
    timeout : BOOL;
END_VAR
VAR
    local_rt : R_TRIG;
    local_rising : BOOL;
    local_prev_phase : INT;
    local_prev_elapsed : INT;
    local_prev_timeout : BOOL;
    local_counted_elapsed : INT;
END_VAR
(* ENGINEERING_CONTRACT
   phase: no-abort start edge -> 1; counted elapsed >= maxDuration -> 3; abort -> 9; otherwise hold 0/1/2/3/9.
   elapsed: +1 only when previous phase 1 or 2, no abort and no start edge; otherwise kept at previous value.
   timeout: set with phase 3 when counted elapsed >= maxDuration; cleared on a no-abort start edge; otherwise held.
   priority: abort > rising start edge > run counting, including same scan start edge.
   start scan does not count. Units: elapsed/maxDuration are scan counts, INT; phase INT 0/1/2/3/9.
   Unspecified: abort plus same-scan start edge keeps phase 9 and consumes that start edge.
*)
(* CONTRACT_RULES [] *)
local_rt(CLK := startBtn);
local_rising := local_rt.Q;

local_prev_phase := phase;
local_prev_elapsed := elapsed;
local_prev_timeout := timeout;

IF abortBtn THEN
    phase := 9;
    elapsed := local_prev_elapsed;
    timeout := local_prev_timeout;
ELSIF local_rising THEN
    phase := 1;
    elapsed := 0;
    timeout := FALSE;
ELSIF (local_prev_phase = 1) OR (local_prev_phase = 2) THEN
    local_counted_elapsed := local_prev_elapsed + 1;
    elapsed := local_counted_elapsed;

    IF local_counted_elapsed >= maxDuration THEN
        timeout := TRUE;
        phase := 3;
    ELSE
        timeout := FALSE;
        IF (local_prev_phase = 2) OR (pv >= setpoint) THEN
            phase := 2;
        ELSE
            phase := 1;
        END_IF;
    END_IF;
ELSE
    phase := local_prev_phase;
    elapsed := local_prev_elapsed;
    timeout := local_prev_timeout;
END_IF;
END_FUNCTION_BLOCK

(* ---- self-hard-02.raw_candidate_01.st ---- *)
FUNCTION_BLOCK FB
VAR_INPUT
    startBtn : BOOL;
    abortBtn : BOOL;
    setpoint : REAL;
    pv : REAL;
    maxDuration : INT;
END_VAR
VAR_OUTPUT
    elapsed : INT;
    phase : INT;
    timeout : BOOL;
END_VAR
VAR
    local_rt : R_TRIG;
    local_rising : BOOL;
    local_prev_phase : INT;
    local_prev_elapsed : INT;
    local_prev_timeout : BOOL;
    local_counted_elapsed : INT;
END_VAR
(* ENGINEERING_CONTRACT
   phase: no-abort start edge -> 1; counted elapsed >= maxDuration -> 3; abort -> 9; otherwise hold 0/1/2/3/9.
   elapsed: +1 only when previous phase 1 or 2, no abort and no start edge; otherwise kept at previous value.
   timeout: set with phase 3 when counted elapsed >= maxDuration; cleared on a no-abort start edge; otherwise held.
   priority: abort > rising start edge > run counting, including same scan start edge.
   start scan does not count. Units: elapsed/maxDuration are scan counts, INT; phase INT 0/1/2/3/9.
   Unspecified: abort plus same-scan start edge keeps phase 9 and consumes that start edge.
*)
(* CONTRACT_RULES [] *)
local_rt(CLK := startBtn);
local_rising := local_rt.Q;

local_prev_phase := phase;
local_prev_elapsed := elapsed;
local_prev_timeout := timeout;

IF abortBtn THEN
    phase := 9;
    elapsed := local_prev_elapsed;
    timeout := local_prev_timeout;
ELSIF local_rising THEN
    phase := 1;
    elapsed := 0;
    timeout := FALSE;
ELSIF (local_prev_phase = 1) OR (local_prev_phase = 2) THEN
    local_counted_elapsed := local_prev_elapsed + 1;
    elapsed := local_counted_elapsed;

    IF local_counted_elapsed >= maxDuration THEN
        timeout := TRUE;
        phase := 3;
    ELSE
        timeout := FALSE;
        IF (local_prev_phase = 2) OR (pv >= setpoint) THEN
            phase := 2;
        ELSE
            phase := 1;
        END_IF;
    END_IF;
ELSE
    phase := local_prev_phase;
    elapsed := local_prev_elapsed;
    timeout := local_prev_timeout;
END_IF;
END_FUNCTION_BLOCK

(* ---- self-hard-03.candidate_01.st ---- *)
(*
ENGINEERING_CONTRACT
Contract basis: PUB001-PUB007 (operation order, outputs, compact buffer); edges per PUB003.
State/output   Activation                            Retention     Reset  Same-scan priority        Bounds
local history  store pushEn/popEn each scan          VAR static    none   edge=signal AND NOT hist  BOOL
count          pop edge accepted first if count>0;    VAR output    none   pop acts before push      INT 0..8
               push edge accepted then if count<8
full/empty     derived from final count               derived       none   after both edge actions   BOOL, count=8/count=0
head           count=0 -> 0 else fifo[1]              derived       none   after final compaction    INT
fifo           pop shifts valid item i+1 to i;        INOUT buffer  none   shift before push append  valid prefix ordered
               accepted push writes fifo[new count]
*)
(* CONTRACT_RULES [] *)
FUNCTION_BLOCK FB
VAR_INPUT
    pushEn : BOOL;
    pushItem : INT;
    popEn : BOOL;
END_VAR
VAR_INOUT
    fifo : ARRAY[1..8] OF INT;
END_VAR
VAR_OUTPUT
    count : INT;
    full : BOOL;
    empty : BOOL;
    head : INT;
END_VAR
VAR
    local_push_history : BOOL;
    local_pop_history : BOOL;
    local_push_rise : BOOL;
    local_pop_rise : BOOL;
    tmp_i : INT;
END_VAR

local_push_rise := pushEn AND NOT local_push_history;
local_pop_rise := popEn AND NOT local_pop_history;

IF local_pop_rise AND (count > 0) THEN
    IF count > 1 THEN
        FOR tmp_i := 1 TO count - 1 BY 1 DO
            fifo[tmp_i] := fifo[tmp_i + 1];
        END_FOR;
    END_IF;
    count := count - 1;
END_IF;

IF local_push_rise THEN
    IF count < 8 THEN
        count := count + 1;
        fifo[count] := pushItem;
    END_IF;
END_IF;

full := (count = 8);
empty := (count = 0);

IF count = 0 THEN
    head := 0;
ELSE
    head := fifo[1];
END_IF;

local_push_history := pushEn;
local_pop_history := popEn;
END_FUNCTION_BLOCK

(* ---- self-hard-03.candidate_02.st ---- *)
(*
ENGINEERING_CONTRACT
Contract basis: PUB001-PUB007 (operation order, outputs, compact buffer); edges per PUB003.
State/output   Activation                            Retention     Reset  Same-scan priority        Bounds
local history  store pushEn/popEn each scan          VAR static    none   edge=signal AND NOT hist  BOOL
count          pop edge accepted first if count>0;    VAR output    none   pop acts before push      INT 0..8
               push edge accepted then if count<8
full/empty     derived from final count               derived       none   after both edge actions   BOOL, count=8/count=0
head           count=0 -> 0 else fifo[1]              derived       none   after final compaction    INT
fifo           pop shifts valid item i+1 to i;        IN_OUT buffer none   shift before push append  valid prefix ordered
               accepted push writes fifo[new count]
*)
(* CONTRACT_RULES [] *)
FUNCTION_BLOCK FB
VAR_INPUT
    pushEn : BOOL;
    pushItem : INT;
    popEn : BOOL;
END_VAR
VAR_IN_OUT
    fifo : ARRAY[1..8] OF INT;
END_VAR
VAR_OUTPUT
    count : INT;
    full : BOOL;
    empty : BOOL;
    head : INT;
END_VAR
VAR
    local_push_history : BOOL;
    local_pop_history : BOOL;
    local_push_rise : BOOL;
    local_pop_rise : BOOL;
    tmp_i : INT;
END_VAR

local_push_rise := pushEn AND NOT local_push_history;
local_pop_rise := popEn AND NOT local_pop_history;

IF local_pop_rise AND (count > 0) THEN
    IF count > 1 THEN
        FOR tmp_i := 1 TO count - 1 BY 1 DO
            fifo[tmp_i] := fifo[tmp_i + 1];
        END_FOR;
    END_IF;
    count := count - 1;
END_IF;

IF local_push_rise THEN
    IF count < 8 THEN
        count := count + 1;
        fifo[count] := pushItem;
    END_IF;
END_IF;

full := (count = 8);
empty := (count = 0);

IF count = 0 THEN
    head := 0;
ELSE
    head := fifo[1];
END_IF;

local_push_history := pushEn;
local_pop_history := popEn;
END_FUNCTION_BLOCK

(* ---- self-hard-03.raw_candidate_01.st ---- *)
(*
ENGINEERING_CONTRACT
Contract basis: PUB001-PUB007 (operation order, outputs, compact buffer); edges per PUB003.
State/output   Activation                            Retention     Reset  Same-scan priority        Bounds
local history  store pushEn/popEn each scan          VAR static    none   edge=signal AND NOT hist  BOOL
count          pop edge accepted first if count>0;    VAR output    none   pop acts before push      INT 0..8
               push edge accepted then if count<8
full/empty     derived from final count               derived       none   after both edge actions   BOOL, count=8/count=0
head           count=0 -> 0 else fifo[1]              derived       none   after final compaction    INT
fifo           pop shifts valid item i+1 to i;        INOUT buffer  none   shift before push append  valid prefix ordered
               accepted push writes fifo[new count]
*)
(* CONTRACT_RULES [] *)
FUNCTION_BLOCK FB
VAR_INPUT
    pushEn : BOOL;
    pushItem : INT;
    popEn : BOOL;
END_VAR
VAR_INOUT
    fifo : ARRAY[1..8] OF INT;
END_VAR
VAR_OUTPUT
    count : INT;
    full : BOOL;
    empty : BOOL;
    head : INT;
END_VAR
VAR
    local_push_history : BOOL;
    local_pop_history : BOOL;
    local_push_rise : BOOL;
    local_pop_rise : BOOL;
    tmp_i : INT;
END_VAR

local_push_rise := pushEn AND NOT local_push_history;
local_pop_rise := popEn AND NOT local_pop_history;

IF local_pop_rise AND (count > 0) THEN
    IF count > 1 THEN
        FOR tmp_i := 1 TO count - 1 BY 1 DO
            fifo[tmp_i] := fifo[tmp_i + 1];
        END_FOR;
    END_IF;
    count := count - 1;
END_IF;

IF local_push_rise THEN
    IF count < 8 THEN
        count := count + 1;
        fifo[count] := pushItem;
    END_IF;
END_IF;

full := (count = 8);
empty := (count = 0);

IF count = 0 THEN
    head := 0;
ELSE
    head := fifo[1];
END_IF;

local_push_history := pushEn;
local_pop_history := popEn;
END_FUNCTION_BLOCK

(* ---- self-hard-03.raw_candidate_02.st ---- *)
(*
ENGINEERING_CONTRACT
Contract basis: PUB001-PUB007 (operation order, outputs, compact buffer); edges per PUB003.
State/output   Activation                            Retention     Reset  Same-scan priority        Bounds
local history  store pushEn/popEn each scan          VAR static    none   edge=signal AND NOT hist  BOOL
count          pop edge accepted first if count>0;    VAR output    none   pop acts before push      INT 0..8
               push edge accepted then if count<8
full/empty     derived from final count               derived       none   after both edge actions   BOOL, count=8/count=0
head           count=0 -> 0 else fifo[1]              derived       none   after final compaction    INT
fifo           pop shifts valid item i+1 to i;        IN_OUT buffer none   shift before push append  valid prefix ordered
               accepted push writes fifo[new count]
*)
(* CONTRACT_RULES [] *)
FUNCTION_BLOCK FB
VAR_INPUT
    pushEn : BOOL;
    pushItem : INT;
    popEn : BOOL;
END_VAR
VAR_IN_OUT
    fifo : ARRAY[1..8] OF INT;
END_VAR
VAR_OUTPUT
    count : INT;
    full : BOOL;
    empty : BOOL;
    head : INT;
END_VAR
VAR
    local_push_history : BOOL;
    local_pop_history : BOOL;
    local_push_rise : BOOL;
    local_pop_rise : BOOL;
    tmp_i : INT;
END_VAR

local_push_rise := pushEn AND NOT local_push_history;
local_pop_rise := popEn AND NOT local_pop_history;

IF local_pop_rise AND (count > 0) THEN
    IF count > 1 THEN
        FOR tmp_i := 1 TO count - 1 BY 1 DO
            fifo[tmp_i] := fifo[tmp_i + 1];
        END_FOR;
    END_IF;
    count := count - 1;
END_IF;

IF local_push_rise THEN
    IF count < 8 THEN
        count := count + 1;
        fifo[count] := pushItem;
    END_IF;
END_IF;

full := (count = 8);
empty := (count = 0);

IF count = 0 THEN
    head := 0;
ELSE
    head := fifo[1];
END_IF;

local_push_history := pushEn;
local_pop_history := popEn;
END_FUNCTION_BLOCK

(* ---- self-hard-04.candidate_01.st ---- *)
FUNCTION_BLOCK FB
(* ENGINEERING_CONTRACT
runningCount: activation=each scan; value=clamp(demand,0,5); reset=none; priority=clamp before pump selection.
leadPump: activation=demand>0 sets initial min or holds; hold=no rotated/insufficient margin; reset=demand<=0 -> 0; change iff rotated AND old-main - min > 50; new lead is used for lag in same scan.
lagPump: activation=demand>=2 on initial, lead-change, or count-rise chooses min non-lead pump; hold=all other demand>=2 scans; reset=demand<=1 -> 0.
units/bounds: demand/pump count 0..5, pump 1..5, runHours LINT hours, hysteresis margin strict >50 h.
*)
(* CONTRACT_RULES [] *)
VAR_INPUT
    demand : INT;
    runHours : ARRAY[1..5] OF LINT;
    rotated : BOOL;
END_VAR
VAR_OUTPUT
    leadPump : INT;
    lagPump : INT;
    runningCount : INT;
END_VAR
VAR
    local_prevLead : INT := 0;
    local_prevCount : INT := 0;
    local_clampedDemand : INT;
    local_minPump : INT;
    local_lagPump : INT;
    local_leadChanged : BOOL;
    local_countRising : BOOL;
    local_index : INT;
END_VAR

    IF demand < 0 THEN
        local_clampedDemand := 0;
    ELSIF demand > 5 THEN
        local_clampedDemand := 5;
    ELSE
        local_clampedDemand := demand;
    END_IF;

    runningCount := local_clampedDemand;
    local_countRising := local_clampedDemand > local_prevCount;

    IF local_clampedDemand = 0 THEN
        leadPump := 0;
        lagPump := 0;
    ELSE
        local_minPump := 1;
        FOR local_index := 2 TO 5 DO
            IF runHours[local_index] < runHours[local_minPump] THEN
                local_minPump := local_index;
            ELSIF runHours[local_index] = runHours[local_minPump] THEN
                IF local_index < local_minPump THEN
                    local_minPump := local_index;
                END_IF;
            END_IF;
        END_FOR;

        IF local_prevLead = 0 THEN
            leadPump := local_minPump;
        ELSE
            leadPump := local_prevLead;
            IF rotated AND (runHours[local_prevLead] - runHours[local_minPump] > 50) THEN
                leadPump := local_minPump;
            END_IF;
        END_IF;

        local_leadChanged := leadPump <> local_prevLead;

        IF local_clampedDemand = 1 THEN
            lagPump := 0;
        ELSE
            IF local_leadChanged OR local_countRising THEN
                local_lagPump := 0;
                FOR local_index := 1 TO 5 DO
                    IF local_index <> leadPump THEN
                        IF local_lagPump = 0 THEN
                            local_lagPump := local_index;
                        ELSIF runHours[local_index] < runHours[local_lagPump] THEN
                            local_lagPump := local_index;
                        ELSIF runHours[local_index] = runHours[local_lagPump] THEN
                            IF local_index < local_lagPump THEN
                                local_lagPump := local_index;
                            END_IF;
                        END_IF;
                    END_IF;
                END_FOR;
                lagPump := local_lagPump;
            END_IF;
        END_IF;
    END_IF;

    local_prevLead := leadPump;
    local_prevCount := runningCount;

END_FUNCTION_BLOCK

(* ---- self-hard-04.raw_candidate_01.st ---- *)
FUNCTION_BLOCK FB
(* ENGINEERING_CONTRACT
runningCount: activation=each scan; value=clamp(demand,0,5); reset=none; priority=clamp before pump selection.
leadPump: activation=demand>0 sets initial min or holds; hold=no rotated/insufficient margin; reset=demand<=0 -> 0; change iff rotated AND old-main - min > 50; new lead is used for lag in same scan.
lagPump: activation=demand>=2 on initial, lead-change, or count-rise chooses min non-lead pump; hold=all other demand>=2 scans; reset=demand<=1 -> 0.
units/bounds: demand/pump count 0..5, pump 1..5, runHours LINT hours, hysteresis margin strict >50 h.
*)
(* CONTRACT_RULES [] *)
VAR_INPUT
    demand : INT;
    runHours : ARRAY[1..5] OF LINT;
    rotated : BOOL;
END_VAR
VAR_OUTPUT
    leadPump : INT;
    lagPump : INT;
    runningCount : INT;
END_VAR
VAR
    local_prevLead : INT := 0;
    local_prevCount : INT := 0;
    local_clampedDemand : INT;
    local_minPump : INT;
    local_lagPump : INT;
    local_leadChanged : BOOL;
    local_countRising : BOOL;
    local_index : INT;
END_VAR

    IF demand < 0 THEN
        local_clampedDemand := 0;
    ELSIF demand > 5 THEN
        local_clampedDemand := 5;
    ELSE
        local_clampedDemand := demand;
    END_IF;

    runningCount := local_clampedDemand;
    local_countRising := local_clampedDemand > local_prevCount;

    IF local_clampedDemand = 0 THEN
        leadPump := 0;
        lagPump := 0;
    ELSE
        local_minPump := 1;
        FOR local_index := 2 TO 5 DO
            IF runHours[local_index] < runHours[local_minPump] THEN
                local_minPump := local_index;
            ELSIF runHours[local_index] = runHours[local_minPump] THEN
                IF local_index < local_minPump THEN
                    local_minPump := local_index;
                END_IF;
            END_IF;
        END_FOR;

        IF local_prevLead = 0 THEN
            leadPump := local_minPump;
        ELSE
            leadPump := local_prevLead;
            IF rotated AND (runHours[local_prevLead] - runHours[local_minPump] > 50) THEN
                leadPump := local_minPump;
            END_IF;
        END_IF;

        local_leadChanged := leadPump <> local_prevLead;

        IF local_clampedDemand = 1 THEN
            lagPump := 0;
        ELSE
            IF local_leadChanged OR local_countRising THEN
                local_lagPump := 0;
                FOR local_index := 1 TO 5 DO
                    IF local_index <> leadPump THEN
                        IF local_lagPump = 0 THEN
                            local_lagPump := local_index;
                        ELSIF runHours[local_index] < runHours[local_lagPump] THEN
                            local_lagPump := local_index;
                        ELSIF runHours[local_index] = runHours[local_lagPump] THEN
                            IF local_index < local_lagPump THEN
                                local_lagPump := local_index;
                            END_IF;
                        END_IF;
                    END_IF;
                END_FOR;
                lagPump := local_lagPump;
            END_IF;
        END_IF;
    END_IF;

    local_prevLead := leadPump;
    local_prevCount := runningCount;

END_FUNCTION_BLOCK

(* ---- self-hard-05.candidate_01.st ---- *)
FUNCTION_BLOCK FB
VAR_INPUT
    runRequest : BOOL;
    flameOK : BOOL;
    o2Valid : BOOL;
    o2PV : REAL;
    baseAir : REAL;
    resetBtn : BOOL;
END_VAR
VAR_OUTPUT
    fuelPermit : BOOL;
    trimEnable : BOOL;
    airTrim : REAL;
    airCommand : REAL;
    tripLatched : BOOL;
    o2Fault : BOOL;
END_VAR
VAR
    tmp_prevReset : BOOL := FALSE;
    tmp_trip : BOOL := FALSE;
    tmp_resetRising : BOOL;
    tmp_rawTrim : REAL;
    tmp_airSum : REAL;
END_VAR

(* ENGINEERING_CONTRACT
   tripLatched: activation runRequest AND NOT flameOK same scan; self-holding;
   reset only rising resetBtn when NOT runRequest AND NOT flameOK; activation wins same-scan reset.
   fuelPermit: runRequest AND flameOK AND NOT tripLatched, not latched.
   o2Fault: NOT o2Valid OR o2PV < 0.0 OR o2PV > 21.0, cuts trim but never fuel.
   trimEnable: fuelPermit AND NOT o2Fault, same scan.
   airTrim: 2.0*(2.0-o2PV), clamp [-10.0,10.0]; zero when trim disabled.
   airCommand: baseAir+airTrim clamp [0.0,100.0]; zero when no fuel permit.
   baseAir itself is unbounded; only final airCommand is bounded. Cite S1-S17/PUB001-PUB065.
*)

(* CONTRACT_RULES [] *)

tmp_resetRising := resetBtn AND NOT tmp_prevReset;

tmp_trip := (runRequest AND NOT flameOK)
            OR (tmp_trip AND NOT (tmp_resetRising AND NOT runRequest AND NOT flameOK));
tripLatched := tmp_trip;
tmp_prevReset := resetBtn;

fuelPermit := runRequest AND flameOK AND NOT tripLatched;

o2Fault := (NOT o2Valid) OR (o2PV < 0.0) OR (o2PV > 21.0);
trimEnable := fuelPermit AND NOT o2Fault;

tmp_rawTrim := 2.0 * (2.0 - o2PV);
IF tmp_rawTrim < -10.0 THEN
    airTrim := -10.0;
ELSIF tmp_rawTrim > 10.0 THEN
    airTrim := 10.0;
ELSE
    airTrim := tmp_rawTrim;
END_IF;

IF NOT trimEnable THEN
    airTrim := 0.0;
END_IF;

IF fuelPermit THEN
    tmp_airSum := baseAir + airTrim;
    IF tmp_airSum < 0.0 THEN
        airCommand := 0.0;
    ELSIF tmp_airSum > 100.0 THEN
        airCommand := 100.0;
    ELSE
        airCommand := tmp_airSum;
    END_IF;
ELSE
    airCommand := 0.0;
END_IF;

END_FUNCTION_BLOCK

(* ---- self-hard-05.raw_candidate_01.st ---- *)
FUNCTION_BLOCK FB
VAR_INPUT
    runRequest : BOOL;
    flameOK : BOOL;
    o2Valid : BOOL;
    o2PV : REAL;
    baseAir : REAL;
    resetBtn : BOOL;
END_VAR
VAR_OUTPUT
    fuelPermit : BOOL;
    trimEnable : BOOL;
    airTrim : REAL;
    airCommand : REAL;
    tripLatched : BOOL;
    o2Fault : BOOL;
END_VAR
VAR
    tmp_prevReset : BOOL := FALSE;
    tmp_trip : BOOL := FALSE;
    tmp_resetRising : BOOL;
    tmp_rawTrim : REAL;
    tmp_airSum : REAL;
END_VAR

(* ENGINEERING_CONTRACT
   tripLatched: activation runRequest AND NOT flameOK same scan; self-holding;
   reset only rising resetBtn when NOT runRequest AND NOT flameOK; activation wins same-scan reset.
   fuelPermit: runRequest AND flameOK AND NOT tripLatched, not latched.
   o2Fault: NOT o2Valid OR o2PV < 0.0 OR o2PV > 21.0, cuts trim but never fuel.
   trimEnable: fuelPermit AND NOT o2Fault, same scan.
   airTrim: 2.0*(2.0-o2PV), clamp [-10.0,10.0]; zero when trim disabled.
   airCommand: baseAir+airTrim clamp [0.0,100.0]; zero when no fuel permit.
   baseAir itself is unbounded; only final airCommand is bounded. Cite S1-S17/PUB001-PUB065.
*)

(* CONTRACT_RULES [] *)

tmp_resetRising := resetBtn AND NOT tmp_prevReset;

tmp_trip := (runRequest AND NOT flameOK)
            OR (tmp_trip AND NOT (tmp_resetRising AND NOT runRequest AND NOT flameOK));
tripLatched := tmp_trip;
tmp_prevReset := resetBtn;

fuelPermit := runRequest AND flameOK AND NOT tripLatched;

o2Fault := (NOT o2Valid) OR (o2PV < 0.0) OR (o2PV > 21.0);
trimEnable := fuelPermit AND NOT o2Fault;

tmp_rawTrim := 2.0 * (2.0 - o2PV);
IF tmp_rawTrim < -10.0 THEN
    airTrim := -10.0;
ELSIF tmp_rawTrim > 10.0 THEN
    airTrim := 10.0;
ELSE
    airTrim := tmp_rawTrim;
END_IF;

IF NOT trimEnable THEN
    airTrim := 0.0;
END_IF;

IF fuelPermit THEN
    tmp_airSum := baseAir + airTrim;
    IF tmp_airSum < 0.0 THEN
        airCommand := 0.0;
    ELSIF tmp_airSum > 100.0 THEN
        airCommand := 100.0;
    ELSE
        airCommand := tmp_airSum;
    END_IF;
ELSE
    airCommand := 0.0;
END_IF;

END_FUNCTION_BLOCK

(* ---- self-hard-06.candidate_01.st ---- *)
FUNCTION_BLOCK FB
VAR_INPUT
    runRequest : BOOL;
    pressure : REAL;
    pressureValid : BOOL;
    fuelFlow : REAL;
    steamFlow : REAL;
    outletCmd : INT;
    outletFeedback : INT;
    resetBtn : BOOL;
END_VAR
VAR_OUTPUT
    tripLatched : BOOL;
    fuelPermit : BOOL;
    currentCauseMask : WORD;
    latchedCauseMask : WORD;
    diagnosticActive : BOOL;
END_VAR
VAR
    local_prevResetBtn : BOOL;
    local_prevTrip : BOOL;
    local_stickCounter : INT;
    local_latchedMask : WORD;
    tmp_resetRising : BOOL;
    tmp_legalReset : BOOL;
    tmp_invalid : BOOL;
    tmp_overpressure : BOOL;
    tmp_tripCondition : BOOL;
    tmp_stickQualified : BOOL;
    tmp_fuelExcess : BOOL;
    tmp_currentMask : WORD;
END_VAR

(* ENGINEERING_CONTRACT
   tripLatched: activate same scan on runRequest AND (NOT pressureValid OR pressure>=4500.0); hold until rising(resetBtn) AND NOT runRequest AND pressureValid AND pressure<=4200.0 [PUB006/PUB007].
   fuelPermit = runRequest AND NOT tripLatched; diagnosticActive iff currentCauseMask<>0 [PUB020].
   currentCauseMask recomputed every scan: 0 when stopped, 1 for invalid data; stick/fuel bits only evaluated during valid overpressure; bit3=8 when no located clue [PUB009-PUB014].
   stick bit1=2 requires three consecutive satisfied scans; any interruption resets count [PUB011/PUB015].
   latchedCauseMask is cumulative bitwise OR of currentCauseMask while tripped, cleared only on legal reset or untripped state [PUB016-PUB018].
   Units: pressure kPa, flows t/h, valve %. Unspecified: scan duration and reset-edge behavior while true trip condition exists.
*)

(* CONTRACT_RULES [] *)

tmp_resetRising := resetBtn AND NOT local_prevResetBtn;
tmp_legalReset := tmp_resetRising AND (NOT runRequest) AND pressureValid AND (pressure <= 4200.0);
tmp_invalid := runRequest AND (NOT pressureValid);
tmp_overpressure := runRequest AND pressureValid AND (pressure >= 4500.0);
tmp_tripCondition := tmp_invalid OR tmp_overpressure;

tripLatched := tmp_tripCondition OR (local_prevTrip AND (NOT tmp_legalReset));

tmp_currentMask := WORD#0;
IF NOT runRequest THEN
    tmp_currentMask := WORD#0;
    local_stickCounter := 0;
ELSIF NOT pressureValid THEN
    tmp_currentMask := WORD#1;
    local_stickCounter := 0;
ELSIF pressure < 4500.0 THEN
    tmp_currentMask := WORD#0;
    local_stickCounter := 0;
ELSE
    tmp_stickQualified := (outletCmd >= 50) AND (outletFeedback <= 10);
    IF tmp_stickQualified THEN
        local_stickCounter := local_stickCounter + 1;
        IF local_stickCounter > 3 THEN
            local_stickCounter := 3;
        END_IF;
    ELSE
        local_stickCounter := 0;
    END_IF;

    IF local_stickCounter >= 3 THEN
        tmp_currentMask := tmp_currentMask OR WORD#2;
    END_IF;

    tmp_fuelExcess := (fuelFlow >= 4.0) AND (steamFlow <= 10.0);
    IF tmp_fuelExcess THEN
        tmp_currentMask := tmp_currentMask OR WORD#4;
    END_IF;

    IF tmp_currentMask = WORD#0 THEN
        tmp_currentMask := WORD#8;
    END_IF;
END_IF;

currentCauseMask := tmp_currentMask;

IF tripLatched THEN
    local_latchedMask := local_latchedMask OR tmp_currentMask;
ELSE
    local_latchedMask := WORD#0;
END_IF;
latchedCauseMask := local_latchedMask;

fuelPermit := runRequest AND NOT tripLatched;
diagnosticActive := (tmp_currentMask <> WORD#0);

local_prevResetBtn := resetBtn;
local_prevTrip := tripLatched;

END_FUNCTION_BLOCK

(* ---- self-hard-06.raw_candidate_01.st ---- *)
FUNCTION_BLOCK FB
VAR_INPUT
    runRequest : BOOL;
    pressure : REAL;
    pressureValid : BOOL;
    fuelFlow : REAL;
    steamFlow : REAL;
    outletCmd : INT;
    outletFeedback : INT;
    resetBtn : BOOL;
END_VAR
VAR_OUTPUT
    tripLatched : BOOL;
    fuelPermit : BOOL;
    currentCauseMask : WORD;
    latchedCauseMask : WORD;
    diagnosticActive : BOOL;
END_VAR
VAR
    local_prevResetBtn : BOOL;
    local_prevTrip : BOOL;
    local_stickCounter : INT;
    local_latchedMask : WORD;
    tmp_resetRising : BOOL;
    tmp_legalReset : BOOL;
    tmp_invalid : BOOL;
    tmp_overpressure : BOOL;
    tmp_tripCondition : BOOL;
    tmp_stickQualified : BOOL;
    tmp_fuelExcess : BOOL;
    tmp_currentMask : WORD;
END_VAR

(* ENGINEERING_CONTRACT
   tripLatched: activate same scan on runRequest AND (NOT pressureValid OR pressure>=4500.0); hold until rising(resetBtn) AND NOT runRequest AND pressureValid AND pressure<=4200.0 [PUB006/PUB007].
   fuelPermit = runRequest AND NOT tripLatched; diagnosticActive iff currentCauseMask<>0 [PUB020].
   currentCauseMask recomputed every scan: 0 when stopped, 1 for invalid data; stick/fuel bits only evaluated during valid overpressure; bit3=8 when no located clue [PUB009-PUB014].
   stick bit1=2 requires three consecutive satisfied scans; any interruption resets count [PUB011/PUB015].
   latchedCauseMask is cumulative bitwise OR of currentCauseMask while tripped, cleared only on legal reset or untripped state [PUB016-PUB018].
   Units: pressure kPa, flows t/h, valve %. Unspecified: scan duration and reset-edge behavior while true trip condition exists.
*)

(* CONTRACT_RULES [] *)

tmp_resetRising := resetBtn AND NOT local_prevResetBtn;
tmp_legalReset := tmp_resetRising AND (NOT runRequest) AND pressureValid AND (pressure <= 4200.0);
tmp_invalid := runRequest AND (NOT pressureValid);
tmp_overpressure := runRequest AND pressureValid AND (pressure >= 4500.0);
tmp_tripCondition := tmp_invalid OR tmp_overpressure;

tripLatched := tmp_tripCondition OR (local_prevTrip AND (NOT tmp_legalReset));

tmp_currentMask := WORD#0;
IF NOT runRequest THEN
    tmp_currentMask := WORD#0;
    local_stickCounter := 0;
ELSIF NOT pressureValid THEN
    tmp_currentMask := WORD#1;
    local_stickCounter := 0;
ELSIF pressure < 4500.0 THEN
    tmp_currentMask := WORD#0;
    local_stickCounter := 0;
ELSE
    tmp_stickQualified := (outletCmd >= 50) AND (outletFeedback <= 10);
    IF tmp_stickQualified THEN
        local_stickCounter := local_stickCounter + 1;
        IF local_stickCounter > 3 THEN
            local_stickCounter := 3;
        END_IF;
    ELSE
        local_stickCounter := 0;
    END_IF;

    IF local_stickCounter >= 3 THEN
        tmp_currentMask := tmp_currentMask OR WORD#2;
    END_IF;

    tmp_fuelExcess := (fuelFlow >= 4.0) AND (steamFlow <= 10.0);
    IF tmp_fuelExcess THEN
        tmp_currentMask := tmp_currentMask OR WORD#4;
    END_IF;

    IF tmp_currentMask = WORD#0 THEN
        tmp_currentMask := WORD#8;
    END_IF;
END_IF;

currentCauseMask := tmp_currentMask;

IF tripLatched THEN
    local_latchedMask := local_latchedMask OR tmp_currentMask;
ELSE
    local_latchedMask := WORD#0;
END_IF;
latchedCauseMask := local_latchedMask;

fuelPermit := runRequest AND NOT tripLatched;
diagnosticActive := (tmp_currentMask <> WORD#0);

local_prevResetBtn := resetBtn;
local_prevTrip := tripLatched;

END_FUNCTION_BLOCK

(* ---- self-medium-01.candidate_01.st ---- *)
TYPE ST_Recipe :
STRUCT
    recipeID : INT;
    totalRatio : REAL;
    temperature : REAL;
END_STRUCT
END_TYPE;

FUNCTION_BLOCK FB
VAR_INPUT
    recipe : ARRAY[1..8] OF ST_Recipe;
    selSlot : INT;
    loadCmd : BOOL;
    running : BOOL;
END_VAR
VAR_OUTPUT
    valid : BOOL;
    loadedID : INT;
END_VAR
VAR
    tmp_prev_load_cmd : BOOL;
END_VAR

(* ENGINEERING_CONTRACT
valid: activates only on an accepted rising loadCmd edge while not running and all checks pass.
valid: holds in every non-accepting scan, including all running scans and held loadCmd.
valid: deactivates on an accepted rising edge when the slot is empty, out of range, or any numeric check fails.
loadedID: updates only on an accepted rising edge; otherwise retains its previous value, including while running.
loadedID: set to recipe[selSlot].recipeID on successful load, or 0 on any accepted invalid load.
Same-scan priority: running suppresses the load-edge action before any slot validation happens.
Boundaries: slots are INT in [1,8]; totalRatio is REAL in [99.0,101.0]; temperature is REAL in [30.0,180.0].
Edge memory: tmp_prev_load_cmd is updated at the end of every scan; no extra reset or interlock is invented.
Initial outputs are unspecified and are left at their default zero values.
*)

(* CONTRACT_RULES [] *)

IF loadCmd AND NOT tmp_prev_load_cmd THEN
    IF NOT running THEN
        IF (selSlot < 1) OR (selSlot > 8) THEN
            valid := FALSE;
            loadedID := 0;
        ELSIF recipe[selSlot].recipeID = 0 THEN
            valid := FALSE;
            loadedID := 0;
        ELSIF (recipe[selSlot].totalRatio < 99.0)
           OR (recipe[selSlot].totalRatio > 101.0) THEN
            valid := FALSE;
            loadedID := 0;
        ELSIF (recipe[selSlot].temperature < 30.0)
           OR (recipe[selSlot].temperature > 180.0) THEN
            valid := FALSE;
            loadedID := 0;
        ELSE
            valid := TRUE;
            loadedID := recipe[selSlot].recipeID;
        END_IF;
    END_IF;
END_IF;

tmp_prev_load_cmd := loadCmd;

END_FUNCTION_BLOCK

(* ---- self-medium-01.raw_candidate_01.st ---- *)
TYPE ST_Recipe :
STRUCT
    recipeID : INT;
    totalRatio : REAL;
    temperature : REAL;
END_STRUCT
END_TYPE

FUNCTION_BLOCK FB
VAR_INPUT
    recipe : ARRAY[1..8] OF ST_Recipe;
    selSlot : INT;
    loadCmd : BOOL;
    running : BOOL;
END_VAR
VAR_OUTPUT
    valid : BOOL;
    loadedID : INT;
END_VAR
VAR
    tmp_prev_load_cmd : BOOL;
END_VAR

(* ENGINEERING_CONTRACT
valid: activates only on an accepted rising loadCmd edge while not running and all checks pass.
valid: holds in every non-accepting scan, including all running scans and held loadCmd.
valid: deactivates on an accepted rising edge when the slot is empty, out of range, or any numeric check fails.
loadedID: updates only on an accepted rising edge; otherwise retains its previous value, including while running.
loadedID: set to recipe[selSlot].recipeID on successful load, or 0 on any accepted invalid load.
Same-scan priority: running suppresses the load-edge action before any slot validation happens.
Boundaries: slots are INT in [1,8]; totalRatio is REAL in [99.0,101.0]; temperature is REAL in [30.0,180.0].
Edge memory: tmp_prev_load_cmd is updated at the end of every scan; no extra reset or interlock is invented.
Initial outputs are unspecified and are left at their default zero values.
*)

(* CONTRACT_RULES [] *)

IF loadCmd AND NOT tmp_prev_load_cmd THEN
    IF NOT running THEN
        IF (selSlot < 1) OR (selSlot > 8) THEN
            valid := FALSE;
            loadedID := 0;
        ELSIF recipe[selSlot].recipeID = 0 THEN
            valid := FALSE;
            loadedID := 0;
        ELSIF (recipe[selSlot].totalRatio < 99.0)
           OR (recipe[selSlot].totalRatio > 101.0) THEN
            valid := FALSE;
            loadedID := 0;
        ELSIF (recipe[selSlot].temperature < 30.0)
           OR (recipe[selSlot].temperature > 180.0) THEN
            valid := FALSE;
            loadedID := 0;
        ELSE
            valid := TRUE;
            loadedID := recipe[selSlot].recipeID;
        END_IF
    END_IF
END_IF

tmp_prev_load_cmd := loadCmd;

END_FUNCTION_BLOCK

(* ---- self-medium-02.candidate_01.st ---- *)
(* ENGINEERING_CONTRACT
 * Activation: enable TRUE -> push rawValue into 8-slot FIFO, then average all currently valid samples.
 * Retention: filteredValue holds its last computed value while enable is FALSE, including persistent disable.
 * Reset: enable FALSE clears ring buffer, count, and write pointer in the same scan; sampleCount := 0 and windowFull := FALSE.
 * Same-scan priority: disabled branch bypasses sampling; count/full reflect end-of-cycle state, filteredValue is not advanced.
 * Bounds/units: sampleCount is INT 0..8, increments each enabled scan until 8 and then stays 8; windowFull is TRUE iff sampleCount = 8.
 *)
(* CONTRACT_RULES [] *)
FUNCTION_BLOCK FB
VAR_INPUT
    enable : BOOL;
    rawValue : REAL;
END_VAR
VAR_OUTPUT
    filteredValue : REAL;
    windowFull : BOOL;
    sampleCount : INT;
END_VAR
VAR
    local_buffer : ARRAY[0..7] OF REAL;
    local_count : INT := 0;
    local_write_index : INT := 0;
    local_sum : REAL := 0.0;
    local_filtered : REAL := 0.0;
    local_i : INT;
END_VAR

IF enable THEN
    local_buffer[local_write_index] := rawValue;
    local_write_index := (local_write_index + 1) MOD 8;

    IF local_count < 8 THEN
        local_count := local_count + 1;
    END_IF;

    local_sum := 0.0;

    IF local_count < 8 THEN
        FOR local_i := 0 TO local_count - 1 DO
            local_sum := local_sum + local_buffer[local_i];
        END_FOR;
        local_filtered := local_sum / INT_TO_REAL(local_count);
    ELSE
        FOR local_i := 0 TO 7 DO
            local_sum := local_sum + local_buffer[local_i];
        END_FOR;
        local_filtered := local_sum / 8.0;
    END_IF;

    sampleCount := local_count;
    windowFull := (local_count = 8);
ELSE
    local_count := 0;
    local_write_index := 0;

    FOR local_i := 0 TO 7 DO
        local_buffer[local_i] := 0.0;
    END_FOR;

    sampleCount := 0;
    windowFull := FALSE;
END_IF;

filteredValue := local_filtered;

END_FUNCTION_BLOCK

(* ---- self-medium-02.raw_candidate_01.st ---- *)
(* ENGINEERING_CONTRACT
 * Activation: enable TRUE -> push rawValue into 8-slot FIFO, then average all currently valid samples.
 * Retention: filteredValue holds its last computed value while enable is FALSE, including persistent disable.
 * Reset: enable FALSE clears ring buffer, count, and write pointer in the same scan; sampleCount := 0 and windowFull := FALSE.
 * Same-scan priority: disabled branch bypasses sampling; count/full reflect end-of-cycle state, filteredValue is not advanced.
 * Bounds/units: sampleCount is INT 0..8, increments each enabled scan until 8 and then stays 8; windowFull is TRUE iff sampleCount = 8.
 *)
(* CONTRACT_RULES [] *)
FUNCTION_BLOCK FB
VAR_INPUT
    enable : BOOL;
    rawValue : REAL;
END_VAR
VAR_OUTPUT
    filteredValue : REAL;
    windowFull : BOOL;
    sampleCount : INT;
END_VAR
VAR
    local_buffer : ARRAY[0..7] OF REAL;
    local_count : INT := 0;
    local_write_index : INT := 0;
    local_sum : REAL := 0.0;
    local_filtered : REAL := 0.0;
    local_i : INT;
END_VAR

IF enable THEN
    local_buffer[local_write_index] := rawValue;
    local_write_index := (local_write_index + 1) MOD 8;

    IF local_count < 8 THEN
        local_count := local_count + 1;
    END_IF;

    local_sum := 0.0;

    IF local_count < 8 THEN
        FOR local_i := 0 TO local_count - 1 DO
            local_sum := local_sum + local_buffer[local_i];
        END_FOR;
        local_filtered := local_sum / INT_TO_REAL(local_count);
    ELSE
        FOR local_i := 0 TO 7 DO
            local_sum := local_sum + local_buffer[local_i];
        END_FOR;
        local_filtered := local_sum / 8.0;
    END_IF;

    sampleCount := local_count;
    windowFull := (local_count = 8);
ELSE
    local_count := 0;
    local_write_index := 0;

    FOR local_i := 0 TO 7 DO
        local_buffer[local_i] := 0.0;
    END_FOR;

    sampleCount := 0;
    windowFull := FALSE;
END_IF;

filteredValue := local_filtered;

END_FUNCTION_BLOCK

(* ---- self-medium-03.candidate_01.st ---- *)
FUNCTION_BLOCK FB
(* ENGINEERING_CONTRACT
   motorUp: IDLE + rising(openBtn) + !closeBtn + !openLimit starts same scan;
   retained in OPENING until openLimit, limit scan returns IDLE and stops same scan.
   motorDown: symmetric with closeBtn/closeLimit.
   errorFlag: any obstacle in any state sets it same scan and stops both directions.
   FAULT retains errorFlag; clear only when !obstacle and rising(openBtn AND closeBtn).
   Reset scan returns IDLE with both motors stopped.
   Priority: obstacle before limit/motion/reset; both buttons pressed together do not start.
*)
(* CONTRACT_RULES [] *)
VAR_INPUT
    openBtn : BOOL;
    closeBtn : BOOL;
    openLimit : BOOL;
    closeLimit : BOOL;
    obstacle : BOOL;
END_VAR
VAR_OUTPUT
    motorUp : BOOL;
    motorDown : BOOL;
    errorFlag : BOOL;
END_VAR
VAR
    state : SINT := 0; (* 0=IDLE, 1=OPENING, 2=CLOSING, 3=FAULT *)
    prevOpenBtn : BOOL := FALSE;
    prevCloseBtn : BOOL := FALSE;
    tmp_risingOpen : BOOL;
    tmp_risingClose : BOOL;
    tmp_risingBoth : BOOL;
END_VAR

motorUp := FALSE;
motorDown := FALSE;
errorFlag := FALSE;

tmp_risingOpen := openBtn AND NOT prevOpenBtn;
tmp_risingClose := closeBtn AND NOT prevCloseBtn;
tmp_risingBoth := openBtn AND closeBtn AND NOT (prevOpenBtn AND prevCloseBtn);

IF obstacle THEN
    errorFlag := TRUE;
    state := 3;
ELSIF state = 3 THEN
    IF tmp_risingBoth THEN
        errorFlag := FALSE;
        state := 0;
    ELSE
        errorFlag := TRUE;
        state := 3;
    END_IF;
ELSIF state = 0 THEN
    IF tmp_risingOpen AND NOT closeBtn AND NOT openLimit THEN
        motorUp := TRUE;
        state := 1;
    ELSIF tmp_risingClose AND NOT openBtn AND NOT closeLimit THEN
        motorDown := TRUE;
        state := 2;
    ELSE
        state := 0;
    END_IF;
ELSIF state = 1 THEN
    IF openLimit THEN
        state := 0;
    ELSE
        motorUp := TRUE;
        state := 1;
    END_IF;
ELSIF state = 2 THEN
    IF closeLimit THEN
        state := 0;
    ELSE
        motorDown := TRUE;
        state := 2;
    END_IF;
END_IF;

prevOpenBtn := openBtn;
prevCloseBtn := closeBtn;
END_FUNCTION_BLOCK

(* ---- self-medium-03.raw_candidate_01.st ---- *)
FUNCTION_BLOCK FB
(* ENGINEERING_CONTRACT
   motorUp: IDLE + rising(openBtn) + !closeBtn + !openLimit starts same scan;
   retained in OPENING until openLimit, limit scan returns IDLE and stops same scan.
   motorDown: symmetric with closeBtn/closeLimit.
   errorFlag: any obstacle in any state sets it same scan and stops both directions.
   FAULT retains errorFlag; clear only when !obstacle and rising(openBtn AND closeBtn).
   Reset scan returns IDLE with both motors stopped.
   Priority: obstacle before limit/motion/reset; both buttons pressed together do not start.
*)
(* CONTRACT_RULES [] *)
VAR_INPUT
    openBtn : BOOL;
    closeBtn : BOOL;
    openLimit : BOOL;
    closeLimit : BOOL;
    obstacle : BOOL;
END_VAR
VAR_OUTPUT
    motorUp : BOOL;
    motorDown : BOOL;
    errorFlag : BOOL;
END_VAR
VAR
    state : SINT := 0; (* 0=IDLE, 1=OPENING, 2=CLOSING, 3=FAULT *)
    prevOpenBtn : BOOL := FALSE;
    prevCloseBtn : BOOL := FALSE;
    tmp_risingOpen : BOOL;
    tmp_risingClose : BOOL;
    tmp_risingBoth : BOOL;
END_VAR

motorUp := FALSE;
motorDown := FALSE;
errorFlag := FALSE;

tmp_risingOpen := openBtn AND NOT prevOpenBtn;
tmp_risingClose := closeBtn AND NOT prevCloseBtn;
tmp_risingBoth := openBtn AND closeBtn AND NOT (prevOpenBtn AND prevCloseBtn);

IF obstacle THEN
    errorFlag := TRUE;
    state := 3;
ELSIF state = 3 THEN
    IF tmp_risingBoth THEN
        errorFlag := FALSE;
        state := 0;
    ELSE
        errorFlag := TRUE;
        state := 3;
    END_IF;
ELSIF state = 0 THEN
    IF tmp_risingOpen AND NOT closeBtn AND NOT openLimit THEN
        motorUp := TRUE;
        state := 1;
    ELSIF tmp_risingClose AND NOT openBtn AND NOT closeLimit THEN
        motorDown := TRUE;
        state := 2;
    ELSE
        state := 0;
    END_IF;
ELSIF state = 1 THEN
    IF openLimit THEN
        state := 0;
    ELSE
        motorUp := TRUE;
        state := 1;
    END_IF;
ELSIF state = 2 THEN
    IF closeLimit THEN
        state := 0;
    ELSE
        motorDown := TRUE;
        state := 2;
    END_IF;
END_IF;

prevOpenBtn := openBtn;
prevCloseBtn := closeBtn;
END_FUNCTION_BLOCK

(* ---- self-medium-04.candidate_01.st ---- *)
FUNCTION_BLOCK FB
VAR_INPUT
    startBtn : BOOL;
    resetBtn : BOOL;
    doneSensor : BOOL;
    targetVol : REAL;
    flowVol : REAL;
END_VAR
VAR_OUTPUT
    valveOpen : BOOL;
    fillsToday : INT;
END_VAR
VAR
    prevStart : BOOL;
    prevReset : BOOL;
    pendingConfirm : BOOL;
    isFilling : BOOL;
    accVolume : REAL;
    tmp_start_edge : BOOL;
    tmp_reset_edge : BOOL;
END_VAR

(* ENGINEERING_CONTRACT
Activation:
- valveOpen opens only on a non-reset start rise from idle/wait-confirm.
- fillsToday increments only after a closed, pending bottle sees doneSensor.
Retention:
- pendingConfirm, isFilling, accVolume and fillsToday persist between scans.
- fillsToday saturates at 32767.
Reset:
- reset rise clears count/volume/pending, closes valve, ignores same-scan start/flow/done.
Same-scan priority:
reset > idle/wait start > flow add and close > done confirmation.
Boundaries:
- volume closes at accVolume >= targetVol; start scan flow is included.
*)

(* CONTRACT_RULES [] *)

tmp_start_edge := startBtn AND NOT prevStart;
tmp_reset_edge := resetBtn AND NOT prevReset;

IF tmp_reset_edge THEN
    fillsToday := 0;
    accVolume := 0.0;
    valveOpen := FALSE;
    pendingConfirm := FALSE;
    isFilling := FALSE;
ELSE
    IF tmp_start_edge AND NOT isFilling THEN
        pendingConfirm := FALSE;
        accVolume := 0.0;
        valveOpen := TRUE;
        isFilling := TRUE;
    END_IF;

    IF isFilling THEN
        accVolume := accVolume + flowVol;
        IF accVolume >= targetVol THEN
            valveOpen := FALSE;
            isFilling := FALSE;
            pendingConfirm := TRUE;
        END_IF;
    END_IF;

    IF pendingConfirm AND doneSensor THEN
        IF fillsToday < 32767 THEN
            fillsToday := fillsToday + 1;
        END_IF;
        pendingConfirm := FALSE;
    END_IF;
END_IF;

prevStart := startBtn;
prevReset := resetBtn;

END_FUNCTION_BLOCK

(* ---- self-medium-04.raw_candidate_01.st ---- *)
FUNCTION_BLOCK FB
VAR_INPUT
    startBtn : BOOL;
    resetBtn : BOOL;
    doneSensor : BOOL;
    targetVol : REAL;
    flowVol : REAL;
END_VAR
VAR_OUTPUT
    valveOpen : BOOL;
    fillsToday : INT;
END_VAR
VAR
    prevStart : BOOL;
    prevReset : BOOL;
    pendingConfirm : BOOL;
    isFilling : BOOL;
    accVolume : REAL;
    tmp_start_edge : BOOL;
    tmp_reset_edge : BOOL;
END_VAR

(* ENGINEERING_CONTRACT
Activation:
- valveOpen opens only on a non-reset start rise from idle/wait-confirm.
- fillsToday increments only after a closed, pending bottle sees doneSensor.
Retention:
- pendingConfirm, isFilling, accVolume and fillsToday persist between scans.
- fillsToday saturates at 32767.
Reset:
- reset rise clears count/volume/pending, closes valve, ignores same-scan start/flow/done.
Same-scan priority:
reset > idle/wait start > flow add and close > done confirmation.
Boundaries:
- volume closes at accVolume >= targetVol; start scan flow is included.
*)

(* CONTRACT_RULES [] *)

tmp_start_edge := startBtn AND NOT prevStart;
tmp_reset_edge := resetBtn AND NOT prevReset;

IF tmp_reset_edge THEN
    fillsToday := 0;
    accVolume := 0.0;
    valveOpen := FALSE;
    pendingConfirm := FALSE;
    isFilling := FALSE;
ELSE
    IF tmp_start_edge AND NOT isFilling THEN
        pendingConfirm := FALSE;
        accVolume := 0.0;
        valveOpen := TRUE;
        isFilling := TRUE;
    END_IF;

    IF isFilling THEN
        accVolume := accVolume + flowVol;
        IF accVolume >= targetVol THEN
            valveOpen := FALSE;
            isFilling := FALSE;
            pendingConfirm := TRUE;
        END_IF;
    END_IF;

    IF pendingConfirm AND doneSensor THEN
        IF fillsToday < 32767 THEN
            fillsToday := fillsToday + 1;
        END_IF;
        pendingConfirm := FALSE;
    END_IF;
END_IF;

prevStart := startBtn;
prevReset := resetBtn;

END_FUNCTION_BLOCK

(* ---- self-medium-05.candidate_01.st ---- *)
FUNCTION_BLOCK FB
VAR_INPUT
    enable : BOOL;
    resetBtn : BOOL;
    scanSeconds : LREAL;
    steamFlow : LREAL;
    fuelFlow : LREAL;
    steamTemp : LREAL;
    steamPressure : LREAL;
END_VAR
VAR_OUTPUT
    qualified : BOOL;
    dataFault : BOOL;
    qualifiedTon : LREAL;
    fuelTon : LREAL;
    revenue : LREAL;
    cost : LREAL;
    netProfit : LREAL;
END_VAR
VAR
    tmp_PrevReset : BOOL := FALSE;
    tmp_RisingReset : BOOL;
END_VAR

(* ENGINEERING_CONTRACT
   qualified: combinational true when steamTemp in [447.0,453.0] AND steamPressure in [3750.0,3850.0], inclusive.
   dataFault: combinational true when scanSeconds<=0.0 or >10.0, steamFlow outside [0.0,90.0], or fuelFlow outside [0.0,6.0].
   qualifiedTon: on reset rising edge -> 0.0 and no accumulation; otherwise add if enable AND !dataFault AND qualified, else hold.
   fuelTon: on reset rising edge -> 0.0 and no accumulation; otherwise add if enable AND !dataFault, else hold.
   revenue, cost, netProfit update every scan from current tonnage; units are t and CNY.
   reset edge has priority over disable and fault; fault flag is still reported.
*)
(* CONTRACT_RULES [] *)

tmp_RisingReset := resetBtn AND NOT tmp_PrevReset;

dataFault := (scanSeconds <= 0.0)
    OR (scanSeconds > 10.0)
    OR (steamFlow < 0.0)
    OR (steamFlow > 90.0)
    OR (fuelFlow < 0.0)
    OR (fuelFlow > 6.0);

qualified := (steamTemp >= 447.0)
    AND (steamTemp <= 453.0)
    AND (steamPressure >= 3750.0)
    AND (steamPressure <= 3850.0);

IF tmp_RisingReset THEN
    qualifiedTon := 0.0;
    fuelTon := 0.0;
ELSE
    IF enable AND NOT dataFault THEN
        fuelTon := fuelTon + fuelFlow * scanSeconds / 1000.0;

        IF qualified THEN
            qualifiedTon := qualifiedTon + steamFlow * scanSeconds / 1000.0;
        END_IF;
    END_IF;
END_IF;

revenue := qualifiedTon * 280.0;
cost := fuelTon * 1500.0;
netProfit := revenue - cost;

tmp_PrevReset := resetBtn;

END_FUNCTION_BLOCK

(* ---- self-medium-05.raw_candidate_01.st ---- *)
FUNCTION_BLOCK FB
VAR_INPUT
    enable : BOOL;
    resetBtn : BOOL;
    scanSeconds : LREAL;
    steamFlow : LREAL;
    fuelFlow : LREAL;
    steamTemp : LREAL;
    steamPressure : LREAL;
END_VAR
VAR_OUTPUT
    qualified : BOOL;
    dataFault : BOOL;
    qualifiedTon : LREAL;
    fuelTon : LREAL;
    revenue : LREAL;
    cost : LREAL;
    netProfit : LREAL;
END_VAR
VAR
    tmp_PrevReset : BOOL := FALSE;
    tmp_RisingReset : BOOL;
END_VAR

(* ENGINEERING_CONTRACT
   qualified: combinational true when steamTemp in [447.0,453.0] AND steamPressure in [3750.0,3850.0], inclusive.
   dataFault: combinational true when scanSeconds<=0.0 or >10.0, steamFlow outside [0.0,90.0], or fuelFlow outside [0.0,6.0].
   qualifiedTon: on reset rising edge -> 0.0 and no accumulation; otherwise add if enable AND !dataFault AND qualified, else hold.
   fuelTon: on reset rising edge -> 0.0 and no accumulation; otherwise add if enable AND !dataFault, else hold.
   revenue, cost, netProfit update every scan from current tonnage; units are t and CNY.
   reset edge has priority over disable and fault; fault flag is still reported.
*)
(* CONTRACT_RULES [] *)

tmp_RisingReset := resetBtn AND NOT tmp_PrevReset;

dataFault := (scanSeconds <= 0.0)
    OR (scanSeconds > 10.0)
    OR (steamFlow < 0.0)
    OR (steamFlow > 90.0)
    OR (fuelFlow < 0.0)
    OR (fuelFlow > 6.0);

qualified := (steamTemp >= 447.0)
    AND (steamTemp <= 453.0)
    AND (steamPressure >= 3750.0)
    AND (steamPressure <= 3850.0);

IF tmp_RisingReset THEN
    qualifiedTon := 0.0;
    fuelTon := 0.0;
ELSE
    IF enable AND NOT dataFault THEN
        fuelTon := fuelTon + fuelFlow * scanSeconds / 1000.0;

        IF qualified THEN
            qualifiedTon := qualifiedTon + steamFlow * scanSeconds / 1000.0;
        END_IF;
    END_IF;
END_IF;

revenue := qualifiedTon * 280.0;
cost := fuelTon * 1500.0;
netProfit := revenue - cost;

tmp_PrevReset := resetBtn;

END_FUNCTION_BLOCK
